screen "P_Slider_1" 1024x768
   Slider "Default" at 10,10 size 60x160; Caption 'SIMATIC'
   TextField "Label_Default" at 10,172 size 68x16; Text 'Default'
   Slider "BackColor" at 80,10 size 60x160; Caption 'SIMATIC'
   TextField "Label_BackColor" at 80,172 size 68x16; Text 'BackColor'
   Slider "BackFillStyle" at 150,10 size 60x160; Caption 'SIMATIC'
   TextField "Label_BackFillStyle" at 150,172 size 68x16; Text 'BackFillStyle'
   Slider "BarBackColor" at 220,10 size 60x160; Caption 'SIMATIC'
   TextField "Label_BarBackColor" at 220,172 size 68x16; Text 'BarBackColor'
   Slider "BarColor" at 290,10 size 60x160; Caption 'SIMATIC'
   TextField "Label_BarColor" at 290,172 size 68x16; Text 'BarColor'
   Slider "BarOrientation" at 360,10 size 60x160; Caption 'SIMATIC'
   TextField "Label_BarOrientation" at 360,172 size 68x16; Text 'BarOrientation'
   Slider "BarOrientation_2" at 430,10 size 60x160; Caption 'SIMATIC'
   TextField "Label_BarOrientation_2" at 430,172 size 68x16; Text 'BarOrientation_2'
   Slider "BarOrientation_3" at 500,10 size 60x160; Caption 'SIMATIC'
   TextField "Label_BarOrientation_3" at 500,172 size 68x16; Text 'BarOrientation_3'
   Slider "BorderBackColor" at 570,10 size 60x160; Caption 'SIMATIC'
   TextField "Label_BorderBackColor" at 570,172 size 68x16; Text 'BorderBackColor'
   Slider "BorderBrightColor3D" at 640,10 size 60x160; Caption 'SIMATIC'
   TextField "Label_BorderBrightColor3D" at 640,172 size 68x16; Text 'BorderBrightColor3D'
   Slider "BorderColor" at 710,10 size 60x160; Caption 'SIMATIC'
   TextField "Label_BorderColor" at 710,172 size 68x16; Text 'BorderColor'
   Slider "BorderInnerStyle3D" at 780,10 size 60x160; Caption 'SIMATIC'
   TextField "Label_BorderInnerStyle3D" at 780,172 size 68x16; Text 'BorderInnerStyle3D'
   Slider "BorderInnerStyle3D_2" at 850,10 size 60x160; Caption 'SIMATIC'
   TextField "Label_BorderInnerStyle3D_2" at 850,172 size 68x16; Text 'BorderInnerStyle3D_2'
   Slider "BorderInnerWidth3D" at 920,10 size 60x160; Caption 'SIMATIC'
   TextField "Label_BorderInnerWidth3D" at 920,172 size 68x16; Text 'BorderInnerWidth3D'
   Slider "BorderOuterStyle3D" at 10,196 size 60x160; Caption 'SIMATIC'
   TextField "Label_BorderOuterStyle3D" at 10,358 size 68x16; Text 'BorderOuterStyle3D'
   Slider "BorderOuterStyle3D_2" at 80,196 size 60x160; Caption 'SIMATIC'
   TextField "Label_BorderOuterStyle3D_2" at 80,358 size 68x16; Text 'BorderOuterStyle3D_2'
   Slider "BorderOuterWidth3D" at 150,196 size 60x160; Caption 'SIMATIC'
   TextField "Label_BorderOuterWidth3D" at 150,358 size 68x16; Text 'BorderOuterWidth3D'
   Slider "BorderShadeColor3D" at 220,196 size 60x160; Caption 'SIMATIC'
   TextField "Label_BorderShadeColor3D" at 220,358 size 68x16; Text 'BorderShadeColor3D'
   Slider "BorderWidth" at 290,196 size 60x160; Caption 'SIMATIC'
   TextField "Label_BorderWidth" at 290,358 size 68x16; Text 'BorderWidth'
   Slider "CornerRadius" at 360,196 size 60x160; Caption 'SIMATIC'
   TextField "Label_CornerRadius" at 360,358 size 68x16; Text 'CornerRadius'
   Slider "EdgeStyle" at 430,196 size 60x160; Caption 'SIMATIC'
   TextField "Label_EdgeStyle" at 430,358 size 68x16; Text 'EdgeStyle'
   Slider "EdgeStyle_2" at 500,196 size 60x160; Caption 'SIMATIC'
   TextField "Label_EdgeStyle_2" at 500,358 size 68x16; Text 'EdgeStyle_2'
   Slider "EdgeStyle_3" at 570,196 size 60x160; Caption 'SIMATIC'
   TextField "Label_EdgeStyle_3" at 570,358 size 68x16; Text 'EdgeStyle_3'
   Slider "EdgeStyle_4" at 640,196 size 60x160; Caption 'SIMATIC'
   TextField "Label_EdgeStyle_4" at 640,358 size 68x16; Text 'EdgeStyle_4'
   Slider "Flashing" at 710,196 size 60x160; Caption 'SIMATIC'
   TextField "Label_Flashing" at 710,358 size 68x16; Text 'Flashing'
   Slider "FocusColor" at 780,196 size 60x160; Caption 'SIMATIC'
   TextField "Label_FocusColor" at 780,358 size 68x16; Text 'FocusColor'
   Slider "FocusWidth" at 850,196 size 60x160; Caption 'SIMATIC'
   TextField "Label_FocusWidth" at 850,358 size 68x16; Text 'FocusWidth'
   Slider "ForeColor" at 920,196 size 60x160; Caption 'SIMATIC'
   TextField "Label_ForeColor" at 920,358 size 68x16; Text 'ForeColor'
   Slider "LabelColor" at 10,382 size 60x160; Caption 'SIMATIC'
   TextField "Label_LabelColor" at 10,544 size 68x16; Text 'LabelColor'
   Slider "MaximumValue" at 80,382 size 60x160; Caption 'SIMATIC'
   TextField "Label_MaximumValue" at 80,544 size 68x16; Text 'MaximumValue'
   Slider "MinimumValue" at 150,382 size 60x160; Caption 'SIMATIC'
   TextField "Label_MinimumValue" at 150,544 size 68x16; Text 'MinimumValue'
   Slider "RangeLower1Color" at 220,382 size 60x160; Caption 'SIMATIC'
   TextField "Label_RangeLower1Color" at 220,544 size 68x16; Text 'RangeLower1Color'
   Slider "RangeLower1Enabled" at 290,382 size 60x160; Caption 'SIMATIC'
   TextField "Label_RangeLower1Enabled" at 290,544 size 68x16; Text 'RangeLower1Enabled'
   Slider "RangeLower2Color" at 360,382 size 60x160; Caption 'SIMATIC'
   TextField "Label_RangeLower2Color" at 360,544 size 68x16; Text 'RangeLower2Color'
   Slider "RangeLower2Enabled" at 430,382 size 60x160; Caption 'SIMATIC'
   TextField "Label_RangeLower2Enabled" at 430,544 size 68x16; Text 'RangeLower2Enabled'
   Slider "RangeNormalColor" at 500,382 size 60x160; Caption 'SIMATIC'
   TextField "Label_RangeNormalColor" at 500,544 size 68x16; Text 'RangeNormalColor'
   Slider "RangeNormalEnabled" at 570,382 size 60x160; Caption 'SIMATIC'
   TextField "Label_RangeNormalEnabled" at 570,544 size 68x16; Text 'RangeNormalEnabled'
   Slider "RangeUpper1Color" at 640,382 size 60x160; Caption 'SIMATIC'
   TextField "Label_RangeUpper1Color" at 640,544 size 68x16; Text 'RangeUpper1Color'
   Slider "RangeUpper1Enabled" at 710,382 size 60x160; Caption 'SIMATIC'
   TextField "Label_RangeUpper1Enabled" at 710,544 size 68x16; Text 'RangeUpper1Enabled'
   Slider "RangeUpper2Color" at 780,382 size 60x160; Caption 'SIMATIC'
   TextField "Label_RangeUpper2Color" at 780,544 size 68x16; Text 'RangeUpper2Color'
   Slider "RangeUpper2Enabled" at 850,382 size 60x160; Caption 'SIMATIC'
   TextField "Label_RangeUpper2Enabled" at 850,544 size 68x16; Text 'RangeUpper2Enabled'
   Slider "ScalePosition" at 920,382 size 60x160; Caption 'SIMATIC'
   TextField "Label_ScalePosition" at 920,544 size 68x16; Text 'ScalePosition'
   Button "Next" at 982,744 size 40x22; TextOff 'Text'
      on Click: ActivateScreen("P_Slider_2", 0)

screen "P_Slider_2" 1024x768
   Slider "ShowBar" at 10,10 size 60x160; Caption 'SIMATIC'
   TextField "Label_ShowBar" at 10,172 size 68x16; Text 'ShowBar'
   Slider "ShowLimitLines" at 80,10 size 60x160; Caption 'SIMATIC'
   TextField "Label_ShowLimitLines" at 80,172 size 68x16; Text 'ShowLimitLines'
   Slider "ShowLimitMarkers" at 150,10 size 60x160; Caption 'SIMATIC'
   TextField "Label_ShowLimitMarkers" at 150,172 size 68x16; Text 'ShowLimitMarkers'
   Slider "ShowLimitRanges" at 220,10 size 60x160; Caption 'SIMATIC'
   TextField "Label_ShowLimitRanges" at 220,172 size 68x16; Text 'ShowLimitRanges'
   Slider "ShowPosition" at 290,10 size 60x160; Caption 'SIMATIC'
   TextField "Label_ShowPosition" at 290,172 size 68x16; Text 'ShowPosition'
   Slider "ShowScale" at 360,10 size 60x160; Caption 'SIMATIC'
   TextField "Label_ShowScale" at 360,172 size 68x16; Text 'ShowScale'
   Slider "ShowThumb" at 430,10 size 60x160; Caption 'SIMATIC'
   TextField "Label_ShowThumb" at 430,172 size 68x16; Text 'ShowThumb'
   Slider "ShowTickLabels" at 500,10 size 60x160; Caption 'SIMATIC'
   TextField "Label_ShowTickLabels" at 500,172 size 68x16; Text 'ShowTickLabels'
   Slider "ShowTicks" at 570,10 size 60x160; Caption 'SIMATIC'
   TextField "Label_ShowTicks" at 570,172 size 68x16; Text 'ShowTicks'
   Slider "ThumbBackColor" at 640,10 size 60x160; Caption 'SIMATIC'
   TextField "Label_ThumbBackColor" at 640,172 size 68x16; Text 'ThumbBackColor'
   Slider "UseDesignColorSchema" at 710,10 size 60x160; Caption 'SIMATIC'
   TextField "Label_UseDesignColorSchema" at 710,172 size 68x16; Text 'UseDesignColorSchema'
   Button "Next" at 982,744 size 40x22; TextOff 'Text'
      on Click: ActivateScreen("P_Gauge_1", 0)

screen "P_Gauge_1" 1024x768
   Gauge "Default" at 10,10 size 150x150; CaptionText 'SIMATIC'
   TextField "Label_Default" at 10,162 size 158x16; Text 'Default'
   Gauge "AngleMax" at 170,10 size 150x150; CaptionText 'SIMATIC'
   TextField "Label_AngleMax" at 170,162 size 158x16; Text 'AngleMax'
   Gauge "AngleMin" at 330,10 size 150x150; CaptionText 'SIMATIC'
   TextField "Label_AngleMin" at 330,162 size 158x16; Text 'AngleMin'
   Gauge "BackColor" at 490,10 size 150x150; CaptionText 'SIMATIC'
   TextField "Label_BackColor" at 490,162 size 158x16; Text 'BackColor'
   Gauge "BackFillStyle" at 650,10 size 150x150; CaptionText 'SIMATIC'
   TextField "Label_BackFillStyle" at 650,162 size 158x16; Text 'BackFillStyle'
   Gauge "BorderBackColor" at 810,10 size 150x150; CaptionText 'SIMATIC'
   TextField "Label_BorderBackColor" at 810,162 size 158x16; Text 'BorderBackColor'
   Gauge "BorderColor" at 10,186 size 150x150; CaptionText 'SIMATIC'
   TextField "Label_BorderColor" at 10,338 size 158x16; Text 'BorderColor'
   Gauge "BorderWidth" at 170,186 size 150x150; CaptionText 'SIMATIC'
   TextField "Label_BorderWidth" at 170,338 size 158x16; Text 'BorderWidth'
   Gauge "CaptionColor" at 330,186 size 150x150; CaptionText 'SIMATIC'
   TextField "Label_CaptionColor" at 330,338 size 158x16; Text 'CaptionColor'
   Gauge "CaptionTop" at 490,186 size 150x150; CaptionText 'SIMATIC'
   TextField "Label_CaptionTop" at 490,338 size 158x16; Text 'CaptionTop'
   Gauge "CenterColor" at 650,186 size 150x150; CaptionText 'SIMATIC'
   TextField "Label_CenterColor" at 650,338 size 158x16; Text 'CenterColor'
   Gauge "CenterSize" at 810,186 size 150x150; CaptionText 'SIMATIC'
   TextField "Label_CenterSize" at 810,338 size 158x16; Text 'CenterSize'
   Gauge "CornerRadius" at 10,362 size 150x150; CaptionText 'SIMATIC'
   TextField "Label_CornerRadius" at 10,514 size 158x16; Text 'CornerRadius'
   Gauge "DialColor" at 170,362 size 150x150; CaptionText 'SIMATIC'
   TextField "Label_DialColor" at 170,514 size 158x16; Text 'DialColor'
   Gauge "DialFillStyle" at 330,362 size 150x150; CaptionText 'SIMATIC'
   TextField "Label_DialFillStyle" at 330,514 size 158x16; Text 'DialFillStyle'
   Gauge "DialSize" at 490,362 size 150x150; CaptionText 'SIMATIC'
   TextField "Label_DialSize" at 490,514 size 158x16; Text 'DialSize'
   Gauge "EdgeStyle" at 650,362 size 150x150; CaptionText 'SIMATIC'
   TextField "Label_EdgeStyle" at 650,514 size 158x16; Text 'EdgeStyle'
   Gauge "EdgeStyle_2" at 810,362 size 150x150; CaptionText 'SIMATIC'
   TextField "Label_EdgeStyle_2" at 810,514 size 158x16; Text 'EdgeStyle_2'
   Gauge "EdgeStyle_3" at 10,538 size 150x150; CaptionText 'SIMATIC'
   TextField "Label_EdgeStyle_3" at 10,690 size 158x16; Text 'EdgeStyle_3'
   Gauge "EdgeStyle_4" at 170,538 size 150x150; CaptionText 'SIMATIC'
   TextField "Label_EdgeStyle_4" at 170,690 size 158x16; Text 'EdgeStyle_4'
   Gauge "Gradation" at 330,538 size 150x150; CaptionText 'SIMATIC'
   TextField "Label_Gradation" at 330,690 size 158x16; Text 'Gradation'
   Gauge "InnerDialColor" at 490,538 size 150x150; CaptionText 'SIMATIC'
   TextField "Label_InnerDialColor" at 490,690 size 158x16; Text 'InnerDialColor'
   Gauge "InnerDialInnerDistance" at 650,538 size 150x150; CaptionText 'SIMATIC'
   TextField "Label_InnerDialInnerDistance" at 650,690 size 158x16; Text 'InnerDialInnerDistance'
   Gauge "InnerDialOuterDistance" at 810,538 size 150x150; CaptionText 'SIMATIC'
   TextField "Label_InnerDialOuterDistance" at 810,690 size 158x16; Text 'InnerDialOuterDistance'
   Button "Next" at 982,744 size 40x22; TextOff 'Text'
      on Click: ActivateScreen("P_Gauge_2", 0)

screen "P_Gauge_2" 1024x768
   Gauge "LockSquaredExtent" at 10,10 size 150x150; CaptionText 'SIMATIC'
   TextField "Label_LockSquaredExtent" at 10,162 size 158x16; Text 'LockSquaredExtent'
   Gauge "MaximumValue" at 170,10 size 150x150; CaptionText 'SIMATIC'
   TextField "Label_MaximumValue" at 170,162 size 158x16; Text 'MaximumValue'
   Gauge "MinimumValue" at 330,10 size 150x150; CaptionText 'SIMATIC'
   TextField "Label_MinimumValue" at 330,162 size 158x16; Text 'MinimumValue'
   Gauge "NeedleHeight" at 490,10 size 150x150; CaptionText 'SIMATIC'
   TextField "Label_NeedleHeight" at 490,162 size 158x16; Text 'NeedleHeight'
   Gauge "PointerColor" at 650,10 size 150x150; CaptionText 'SIMATIC'
   TextField "Label_PointerColor" at 650,162 size 158x16; Text 'PointerColor'
   Gauge "RangeLower1Color" at 810,10 size 150x150; CaptionText 'SIMATIC'
   TextField "Label_RangeLower1Color" at 810,162 size 158x16; Text 'RangeLower1Color'
   Gauge "RangeLower1Enabled" at 10,186 size 150x150; CaptionText 'SIMATIC'
   TextField "Label_RangeLower1Enabled" at 10,338 size 158x16; Text 'RangeLower1Enabled'
   Gauge "RangeLower2Color" at 170,186 size 150x150; CaptionText 'SIMATIC'
   TextField "Label_RangeLower2Color" at 170,338 size 158x16; Text 'RangeLower2Color'
   Gauge "RangeLower2Enabled" at 330,186 size 150x150; CaptionText 'SIMATIC'
   TextField "Label_RangeLower2Enabled" at 330,338 size 158x16; Text 'RangeLower2Enabled'
   Gauge "RangeNormalColor" at 490,186 size 150x150; CaptionText 'SIMATIC'
   TextField "Label_RangeNormalColor" at 490,338 size 158x16; Text 'RangeNormalColor'
   Gauge "RangeNormalEnabled" at 650,186 size 150x150; CaptionText 'SIMATIC'
   TextField "Label_RangeNormalEnabled" at 650,338 size 158x16; Text 'RangeNormalEnabled'
   Gauge "RangeUpper1Color" at 810,186 size 150x150; CaptionText 'SIMATIC'
   TextField "Label_RangeUpper1Color" at 810,338 size 158x16; Text 'RangeUpper1Color'
   Gauge "RangeUpper1Enabled" at 10,362 size 150x150; CaptionText 'SIMATIC'
   TextField "Label_RangeUpper1Enabled" at 10,514 size 158x16; Text 'RangeUpper1Enabled'
   Gauge "RangeUpper1Start" at 170,362 size 150x150; CaptionText 'SIMATIC'
   TextField "Label_RangeUpper1Start" at 170,514 size 158x16; Text 'RangeUpper1Start'
   Gauge "RangeUpper2Color" at 330,362 size 150x150; CaptionText 'SIMATIC'
   TextField "Label_RangeUpper2Color" at 330,514 size 158x16; Text 'RangeUpper2Color'
   Gauge "RangeUpper2Enabled" at 490,362 size 150x150; CaptionText 'SIMATIC'
   TextField "Label_RangeUpper2Enabled" at 490,514 size 158x16; Text 'RangeUpper2Enabled'
   Gauge "RangeUpper2Start" at 650,362 size 150x150; CaptionText 'SIMATIC'
   TextField "Label_RangeUpper2Start" at 650,514 size 158x16; Text 'RangeUpper2Start'
   Gauge "ScaleLabelColor" at 810,362 size 150x150; CaptionText 'SIMATIC'
   TextField "Label_ScaleLabelColor" at 810,514 size 158x16; Text 'ScaleLabelColor'
   Gauge "ScaleTickColor" at 10,538 size 150x150; CaptionText 'SIMATIC'
   TextField "Label_ScaleTickColor" at 10,690 size 158x16; Text 'ScaleTickColor'
   Gauge "ScaleTickLabelPosition" at 170,538 size 150x150; CaptionText 'SIMATIC'
   TextField "Label_ScaleTickLabelPosition" at 170,690 size 158x16; Text 'ScaleTickLabelPosition'
   Gauge "ScaleTickLength" at 330,538 size 150x150; CaptionText 'SIMATIC'
   TextField "Label_ScaleTickLength" at 330,690 size 158x16; Text 'ScaleTickLength'
   Gauge "ScaleTickPosition" at 490,538 size 150x150; CaptionText 'SIMATIC'
   TextField "Label_ScaleTickPosition" at 490,690 size 158x16; Text 'ScaleTickPosition'
   Gauge "ShowDecimalPoint" at 650,538 size 150x150; CaptionText 'SIMATIC'
   TextField "Label_ShowDecimalPoint" at 650,690 size 158x16; Text 'ShowDecimalPoint'
   Gauge "ShowInnerDial" at 810,538 size 150x150; CaptionText 'SIMATIC'
   TextField "Label_ShowInnerDial" at 810,690 size 158x16; Text 'ShowInnerDial'
   Button "Next" at 982,744 size 40x22; TextOff 'Text'
      on Click: ActivateScreen("P_Gauge_3", 0)

screen "P_Gauge_3" 1024x768
   Gauge "ShowLimitRanges" at 10,10 size 150x150; CaptionText 'SIMATIC'
   TextField "Label_ShowLimitRanges" at 10,162 size 158x16; Text 'ShowLimitRanges'
   Gauge "ShowPeakValuePointer" at 170,10 size 150x150; CaptionText 'SIMATIC'
   TextField "Label_ShowPeakValuePointer" at 170,162 size 158x16; Text 'ShowPeakValuePointer'
   Gauge "UnitColor" at 330,10 size 150x150; CaptionText 'SIMATIC'
   TextField "Label_UnitColor" at 330,162 size 158x16; Text 'UnitColor'
   Gauge "UnitTop" at 490,10 size 150x150; CaptionText 'SIMATIC'
   TextField "Label_UnitTop" at 490,162 size 158x16; Text 'UnitTop'
   Gauge "UseDesignColorSchema" at 650,10 size 150x150; CaptionText 'SIMATIC'
   TextField "Label_UseDesignColorSchema" at 650,162 size 158x16; Text 'UseDesignColorSchema'
   Button "Next" at 982,744 size 40x22; TextOff 'Text'
      on Click: ActivateScreen("P_Clock_1", 0)

screen "P_Clock_1" 1024x768
   Clock "Default" at 10,10 size 150x150
   TextField "Label_Default" at 10,162 size 158x16; Text 'Default'
   Clock "Analog" at 170,10 size 150x150
   TextField "Label_Analog" at 170,162 size 158x16; Text 'Analog'
   Clock "BackFillStyle" at 330,10 size 150x150
   TextField "Label_BackFillStyle" at 330,162 size 158x16; Text 'BackFillStyle'
   Clock "BorderBackColor" at 490,10 size 150x150
   TextField "Label_BorderBackColor" at 490,162 size 158x16; Text 'BorderBackColor'
   Clock "BorderColor" at 650,10 size 150x150
   TextField "Label_BorderColor" at 650,162 size 158x16; Text 'BorderColor'
   Clock "BorderWidth" at 810,10 size 150x150
   TextField "Label_BorderWidth" at 810,162 size 158x16; Text 'BorderWidth'
   Clock "CornerRadius" at 10,186 size 150x150
   TextField "Label_CornerRadius" at 10,338 size 158x16; Text 'CornerRadius'
   Clock "DialColor" at 170,186 size 150x150
   TextField "Label_DialColor" at 170,338 size 158x16; Text 'DialColor'
   Clock "EdgeStyle" at 330,186 size 150x150
   TextField "Label_EdgeStyle" at 330,338 size 158x16; Text 'EdgeStyle'
   Clock "EdgeStyle_2" at 490,186 size 150x150
   TextField "Label_EdgeStyle_2" at 490,338 size 158x16; Text 'EdgeStyle_2'
   Clock "EdgeStyle_3" at 650,186 size 150x150
   TextField "Label_EdgeStyle_3" at 650,338 size 158x16; Text 'EdgeStyle_3'
   Clock "EdgeStyle_4" at 810,186 size 150x150
   TextField "Label_EdgeStyle_4" at 810,338 size 158x16; Text 'EdgeStyle_4'
   Clock "Flashing" at 10,362 size 150x150
   TextField "Label_Flashing" at 10,514 size 158x16; Text 'Flashing'
   Clock "HourNeedleHeight" at 170,362 size 150x150
   TextField "Label_HourNeedleHeight" at 170,514 size 158x16; Text 'HourNeedleHeight'
   Clock "HourNeedleWidth" at 330,362 size 150x150
   TextField "Label_HourNeedleWidth" at 330,514 size 158x16; Text 'HourNeedleWidth'
   Clock "LockSquaredExtent" at 490,362 size 150x150
   TextField "Label_LockSquaredExtent" at 490,514 size 158x16; Text 'LockSquaredExtent'
   Clock "MinuteNeedleHeight" at 650,362 size 150x150
   TextField "Label_MinuteNeedleHeight" at 650,514 size 158x16; Text 'MinuteNeedleHeight'
   Clock "MinuteNeedleWidth" at 810,362 size 150x150
   TextField "Label_MinuteNeedleWidth" at 810,514 size 158x16; Text 'MinuteNeedleWidth'
   Clock "NeedleBorderColor" at 10,538 size 150x150
   TextField "Label_NeedleBorderColor" at 10,690 size 158x16; Text 'NeedleBorderColor'
   Clock "NeedleColor" at 170,538 size 150x150
   TextField "Label_NeedleColor" at 170,690 size 158x16; Text 'NeedleColor'
   Clock "NeedleFillStyle" at 330,538 size 150x150
   TextField "Label_NeedleFillStyle" at 330,690 size 158x16; Text 'NeedleFillStyle'
   Clock "NumberStyle" at 490,538 size 150x150
   TextField "Label_NumberStyle" at 490,690 size 158x16; Text 'NumberStyle'
   Clock "NumberStyle_2" at 650,538 size 150x150
   TextField "Label_NumberStyle_2" at 650,690 size 158x16; Text 'NumberStyle_2'
   Clock "SecondNeedleHeight" at 810,538 size 150x150
   TextField "Label_SecondNeedleHeight" at 810,690 size 158x16; Text 'SecondNeedleHeight'
   Button "Next" at 982,744 size 40x22; TextOff 'Text'
      on Click: ActivateScreen("P_Clock_2", 0)

screen "P_Clock_2" 1024x768
   Clock "SecondNeedleWidth" at 10,10 size 150x150
   TextField "Label_SecondNeedleWidth" at 10,162 size 158x16; Text 'SecondNeedleWidth'
   Clock "ShowTicks" at 170,10 size 150x150
   TextField "Label_ShowTicks" at 170,162 size 158x16; Text 'ShowTicks'
   Clock "TickDistance" at 330,10 size 150x150
   TextField "Label_TickDistance" at 330,162 size 158x16; Text 'TickDistance'
   Clock "TickStyle" at 490,10 size 150x150
   TextField "Label_TickStyle" at 490,162 size 158x16; Text 'TickStyle'
   Clock "TicksColor" at 650,10 size 150x150
   TextField "Label_TicksColor" at 650,162 size 158x16; Text 'TicksColor'
   Clock "UseDesignColorSchema" at 810,10 size 150x150
   TextField "Label_UseDesignColorSchema" at 810,162 size 158x16; Text 'UseDesignColorSchema'
   Button "Next" at 982,744 size 40x22; TextOff 'Text'
      on Click: ActivateScreen("P_Line_1", 0)

screen "P_IOField_1" 1024x768
   IOField "Default" at 10,10 size 100x30
   TextField "Label_Default" at 10,42 size 108x16; Text 'Default'
   IOField "AboveUpperLimitColor" at 120,10 size 100x30
   TextField "Label_AboveUpperLimitColor" at 120,42 size 108x16; Text 'AboveUpperLimitColor'
   IOField "BackColor" at 230,10 size 100x30
   TextField "Label_BackColor" at 230,42 size 108x16; Text 'BackColor'
   IOField "BackFillStyle" at 340,10 size 100x30
   TextField "Label_BackFillStyle" at 340,42 size 108x16; Text 'BackFillStyle'
   IOField "BelowLowerLimitColor" at 450,10 size 100x30
   TextField "Label_BelowLowerLimitColor" at 450,42 size 108x16; Text 'BelowLowerLimitColor'
   IOField "BorderBackColor" at 560,10 size 100x30
   TextField "Label_BorderBackColor" at 560,42 size 108x16; Text 'BorderBackColor'
   IOField "BorderColor" at 670,10 size 100x30
   TextField "Label_BorderColor" at 670,42 size 108x16; Text 'BorderColor'
   IOField "BorderWidth" at 780,10 size 100x30
   TextField "Label_BorderWidth" at 780,42 size 108x16; Text 'BorderWidth'
   IOField "BottomMargin" at 890,10 size 100x30
   TextField "Label_BottomMargin" at 890,42 size 108x16; Text 'BottomMargin'
   IOField "CornerRadius" at 10,66 size 100x30
   TextField "Label_CornerRadius" at 10,98 size 108x16; Text 'CornerRadius'
   IOField "DataFormat_3" at 120,66 size 100x30
   TextField "Label_DataFormat_3" at 120,98 size 108x16; Text 'DataFormat_3'
   IOField "EdgeStyle" at 230,66 size 100x30
   TextField "Label_EdgeStyle" at 230,98 size 108x16; Text 'EdgeStyle'
   IOField "EdgeStyle_2" at 340,66 size 100x30
   TextField "Label_EdgeStyle_2" at 340,98 size 108x16; Text 'EdgeStyle_2'
   IOField "EdgeStyle_3" at 450,66 size 100x30
   TextField "Label_EdgeStyle_3" at 450,98 size 108x16; Text 'EdgeStyle_3'
   IOField "EdgeStyle_4" at 560,66 size 100x30
   TextField "Label_EdgeStyle_4" at 560,98 size 108x16; Text 'EdgeStyle_4'
   IOField "FieldLength" at 670,66 size 100x30
   TextField "Label_FieldLength" at 670,98 size 108x16; Text 'FieldLength'
   IOField "FitToLargest" at 780,66 size 100x30
   TextField "Label_FitToLargest" at 780,98 size 108x16; Text 'FitToLargest'
   IOField "Flashing" at 890,66 size 100x30
   TextField "Label_Flashing" at 890,98 size 108x16; Text 'Flashing'
   IOField "ForeColor" at 10,122 size 100x30
   TextField "Label_ForeColor" at 10,154 size 108x16; Text 'ForeColor'
   IOField "FormatPattern" at 120,122 size 100x30; FormatPattern 99.9
   TextField "Label_FormatPattern" at 120,154 size 108x16; Text 'FormatPattern'
   IOField "HorizontalAlignment" at 230,122 size 100x30
   TextField "Label_HorizontalAlignment" at 230,154 size 108x16; Text 'HorizontalAlignment'
   IOField "HorizontalAlignment_2" at 340,122 size 100x30
   TextField "Label_HorizontalAlignment_2" at 340,154 size 108x16; Text 'HorizontalAlignment_2'
   IOField "LeftMargin" at 450,122 size 100x30
   TextField "Label_LeftMargin" at 450,154 size 108x16; Text 'LeftMargin'
   IOField "Mode" at 560,122 size 100x30
   TextField "Label_Mode" at 560,154 size 108x16; Text 'Mode'
   IOField "Mode_2" at 670,122 size 100x30
   TextField "Label_Mode_2" at 670,154 size 108x16; Text 'Mode_2'
   IOField "RightMargin" at 780,122 size 100x30
   TextField "Label_RightMargin" at 780,154 size 108x16; Text 'RightMargin'
   IOField "ShiftDecimalPoint" at 890,122 size 100x30
   TextField "Label_ShiftDecimalPoint" at 890,154 size 108x16; Text 'ShiftDecimalPoint'
   IOField "ShowLeadingZeros" at 10,178 size 100x30
   TextField "Label_ShowLeadingZeros" at 10,210 size 108x16; Text 'ShowLeadingZeros'
   IOField "TopMargin" at 120,178 size 100x30
   TextField "Label_TopMargin" at 120,210 size 108x16; Text 'TopMargin'
   IOField "Unit" at 230,178 size 100x30; Unit mm
   TextField "Label_Unit" at 230,210 size 108x16; Text 'Unit'
   IOField "UseDesignColorSchema" at 340,178 size 100x30
   TextField "Label_UseDesignColorSchema" at 340,210 size 108x16; Text 'UseDesignColorSchema'
   IOField "VerticalAlignment" at 450,178 size 100x30
   TextField "Label_VerticalAlignment" at 450,210 size 108x16; Text 'VerticalAlignment'
   IOField "VerticalAlignment_2" at 560,178 size 100x30
   TextField "Label_VerticalAlignment_2" at 560,210 size 108x16; Text 'VerticalAlignment_2'
   Button "Next" at 982,744 size 40x22; TextOff 'Text'
      on Click: ActivateScreen("P_Button_1", 0)

screen "D_Bar_1" 1024x768
   Bar "Static" at 6,4 size 40x120
   TextField "Label_Static" at 6,156 size 88x16; Text 'Static'
   Bar "A_Range" at 98,4 size 40x120
      Appearance <- "D_Range"
   TextField "Label_A_Range" at 98,156 size 88x16; Text 'A_Range'
   Bar "A_Flash" at 190,4 size 40x120
      Appearance <- "D_Range"
   TextField "Label_A_Flash" at 190,156 size 88x16; Text 'A_Flash'
   Bar "A_Bit" at 282,4 size 40x120
      Appearance <- "D_Bool"
   TextField "Label_A_Bit" at 282,156 size 88x16; Text 'A_Bit'
   Bar "A_Bits" at 374,4 size 40x120
      Appearance <- "D_Bits"
   TextField "Label_A_Bits" at 374,156 size 88x16; Text 'A_Bits'
   Bar "V_Range" at 466,4 size 40x120
      Visibility <- "D_Range"
   TextField "Label_V_Range" at 466,156 size 88x16; Text 'V_Range'
   Bar "V_Bit" at 558,4 size 40x120
      Visibility <- "D_Vis"
   TextField "Label_V_Bit" at 558,156 size 88x16; Text 'V_Bit'
   Bar "M_H" at 650,4 size 40x120
      HorizontalMovement <- "D_Pct"
   TextField "Label_M_H" at 650,156 size 88x16; Text 'M_H'
   Bar "M_V" at 742,4 size 40x120
      VerticalMovement <- "D_Pct"
   TextField "Label_M_V" at 742,156 size 88x16; Text 'M_V'
   Bar "M_D" at 834,4 size 40x120
      DiagonalMovement <- "D_Pct"
   TextField "Label_M_D" at 834,156 size 88x16; Text 'M_D'
   Bar "M_Direct" at 926,4 size 40x120
      DirectMovement <- "D_X"
      DirectMovement <- "D_Y"
   TextField "Label_M_Direct" at 926,156 size 88x16; Text 'M_Direct'
   Bar "E_Range" at 6,176 size 40x120
      ObjectEnable <- "D_Range"
   TextField "Label_E_Range" at 6,328 size 88x16; Text 'E_Range'
   Bar "E_Bit" at 98,176 size 40x120
      ObjectEnable <- "D_En"
   TextField "Label_E_Bit" at 98,328 size 88x16; Text 'E_Bit'
   Bar "PV_Pct" at 190,176 size 40x120
      ProcessValue <- "D_Pct"
   TextField "Label_PV_Pct" at 190,328 size 88x16; Text 'PV_Pct'
   Bar "PV_Real" at 282,176 size 40x120
      ProcessValue <- "D_Real"
   TextField "Label_PV_Real" at 282,328 size 88x16; Text 'PV_Real'
   Bar "PV_BarR" at 374,176 size 40x120
      ProcessValue <- "D_BarR"
   TextField "Label_PV_BarR" at 374,328 size 88x16; Text 'PV_BarR'
   Bar "PV_Pct_0_100" at 466,176 size 40x120; MinimumValue 0; MaximumValue 100
      ProcessValue <- "D_Pct"
   TextField "Label_PV_Pct_0_100" at 466,328 size 88x16; Text 'PV_Pct_0_100'
   Bar "PV_Pct_MaxMin" at 558,176 size 40x120
      ProcessValue <- "D_Pct"
      MaximumValue <- "D_Max"
      MinimumValue <- "D_Min"
   TextField "Label_PV_Pct_MaxMin" at 558,328 size 88x16; Text 'PV_Pct_MaxMin'
   IOField "State" at 4,742 size 60x22; FormatPattern 9
      ProcessValue <- "D_State"
   Button "S1" at 70,742 size 40x22; TextOff 'S1'
      on Click: "SetS1"()
   Button "S2" at 114,742 size 40x22; TextOff 'S2'
      on Click: "SetS2"()
   Button "S3" at 158,742 size 40x22; TextOff 'S3'
      on Click: "SetS3"()
   Button "S4" at 202,742 size 40x22; TextOff 'S4'
      on Click: "SetS4"()
   Button "Next" at 980,742 size 40x22; TextOff 'Next'
      on Click: ActivateScreen("D_Switch_1", 0)

screen "D_Button_1" 1024x768
   Button "Static" at 6,4 size 100x40; TextOff 'Text'
   TextField "Label_Static" at 6,76 size 148x16; Text 'Static'
   Button "A_Range" at 158,4 size 100x40; TextOff 'Text'
      Appearance <- "D_Range"
   TextField "Label_A_Range" at 158,76 size 148x16; Text 'A_Range'
   Button "A_Flash" at 310,4 size 100x40; TextOff 'Text'
      Appearance <- "D_Range"
   TextField "Label_A_Flash" at 310,76 size 148x16; Text 'A_Flash'
   Button "A_Bit" at 462,4 size 100x40; TextOff 'Text'
      Appearance <- "D_Bool"
   TextField "Label_A_Bit" at 462,76 size 148x16; Text 'A_Bit'
   Button "A_Bits" at 614,4 size 100x40; TextOff 'Text'
      Appearance <- "D_Bits"
   TextField "Label_A_Bits" at 614,76 size 148x16; Text 'A_Bits'
   Button "V_Range" at 766,4 size 100x40; TextOff 'Text'
      Visibility <- "D_Range"
   TextField "Label_V_Range" at 766,76 size 148x16; Text 'V_Range'
   Button "V_Bit" at 6,96 size 100x40; TextOff 'Text'
      Visibility <- "D_Vis"
   TextField "Label_V_Bit" at 6,168 size 148x16; Text 'V_Bit'
   Button "M_H" at 158,96 size 100x40; TextOff 'Text'
      HorizontalMovement <- "D_Pct"
   TextField "Label_M_H" at 158,168 size 148x16; Text 'M_H'
   Button "M_V" at 310,96 size 100x40; TextOff 'Text'
      VerticalMovement <- "D_Pct"
   TextField "Label_M_V" at 310,168 size 148x16; Text 'M_V'
   Button "M_D" at 462,96 size 100x40; TextOff 'Text'
      DiagonalMovement <- "D_Pct"
   TextField "Label_M_D" at 462,168 size 148x16; Text 'M_D'
   Button "M_Direct" at 614,96 size 100x40; TextOff 'Text'
      DirectMovement <- "D_X"
      DirectMovement <- "D_Y"
   TextField "Label_M_Direct" at 614,168 size 148x16; Text 'M_Direct'
   Button "E_Range" at 766,96 size 100x40; TextOff 'Text'
      ObjectEnable <- "D_Range"
   TextField "Label_E_Range" at 766,168 size 148x16; Text 'E_Range'
   Button "E_Bit" at 6,188 size 100x40; TextOff 'Text'
      ObjectEnable <- "D_En"
   TextField "Label_E_Bit" at 6,260 size 148x16; Text 'E_Bit'
   IOField "State" at 4,742 size 60x22; FormatPattern 9
      ProcessValue <- "D_State"
   Button "S1" at 70,742 size 40x22; TextOff 'S1'
      on Click: "SetS1"()
   Button "S2" at 114,742 size 40x22; TextOff 'S2'
      on Click: "SetS2"()
   Button "S3" at 158,742 size 40x22; TextOff 'S3'
      on Click: "SetS3"()
   Button "S4" at 202,742 size 40x22; TextOff 'S4'
      on Click: "SetS4"()
   Button "Next" at 980,742 size 40x22; TextOff 'Next'
      on Click: ActivateScreen("D_SymbolicIOField_1", 0)

screen "D_Circle_1" 1024x768
   TextField "Label_Static" at 6,86 size 98x16; Text 'Static'
   Circle "A_Range" at 108,4 size 50x50
      Appearance <- "D_Range"
   TextField "Label_A_Range" at 108,86 size 98x16; Text 'A_Range'
   Circle "A_Flash" at 210,4 size 50x50
      Appearance <- "D_Range"
   TextField "Label_A_Flash" at 210,86 size 98x16; Text 'A_Flash'
   Circle "A_Bit" at 312,4 size 50x50
      Appearance <- "D_Bool"
   TextField "Label_A_Bit" at 312,86 size 98x16; Text 'A_Bit'
   Circle "A_Bits" at 414,4 size 50x50
      Appearance <- "D_Bits"
   TextField "Label_A_Bits" at 414,86 size 98x16; Text 'A_Bits'
   Circle "V_Range" at 516,4 size 50x50
      Visibility <- "D_Range"
   TextField "Label_V_Range" at 516,86 size 98x16; Text 'V_Range'
   Circle "V_Bit" at 618,4 size 50x50
      Visibility <- "D_Vis"
   TextField "Label_V_Bit" at 618,86 size 98x16; Text 'V_Bit'
   Circle "M_H" at 720,4 size 50x50
      HorizontalMovement <- "D_Pct"
   TextField "Label_M_H" at 720,86 size 98x16; Text 'M_H'
   Circle "M_V" at 822,4 size 50x50
      VerticalMovement <- "D_Pct"
   TextField "Label_M_V" at 822,86 size 98x16; Text 'M_V'
   Circle "M_D" at 6,106 size 50x50
      DiagonalMovement <- "D_Pct"
   TextField "Label_M_D" at 6,188 size 98x16; Text 'M_D'
   Circle "M_Direct" at 108,106 size 50x50
      DirectMovement <- "D_X"
      DirectMovement <- "D_Y"
   TextField "Label_M_Direct" at 108,188 size 98x16; Text 'M_Direct'
   Circle "E_Range" at 210,106 size 50x50
      ObjectEnable <- "D_Range"
   TextField "Label_E_Range" at 210,188 size 98x16; Text 'E_Range'
   Circle "E_Bit" at 312,106 size 50x50
      ObjectEnable <- "D_En"
   TextField "Label_E_Bit" at 312,188 size 98x16; Text 'E_Bit'
   IOField "State" at 4,742 size 60x22; FormatPattern 9
      ProcessValue <- "D_State"
   Button "S1" at 70,742 size 40x22; TextOff 'S1'
      on Click: "SetS1"()
   Button "S2" at 114,742 size 40x22; TextOff 'S2'
      on Click: "SetS2"()
   Button "S3" at 158,742 size 40x22; TextOff 'S3'
      on Click: "SetS3"()
   Button "S4" at 202,742 size 40x22; TextOff 'S4'
      on Click: "SetS4"()
   Button "Next" at 980,742 size 40x22; TextOff 'Next'
      on Click: ActivateScreen("D_Rectangle_1", 0)

screen "D_Clock_1" 1024x768
   Clock "Static" at 6,4 size 150x150
   TextField "Label_Static" at 6,186 size 198x16; Text 'Static'
   Clock "A_Range" at 208,4 size 150x150
      Appearance <- "D_Range"
   TextField "Label_A_Range" at 208,186 size 198x16; Text 'A_Range'
   Clock "A_Flash" at 410,4 size 150x150
      Appearance <- "D_Range"
   TextField "Label_A_Flash" at 410,186 size 198x16; Text 'A_Flash'
   Clock "A_Bit" at 612,4 size 150x150
      Appearance <- "D_Bool"
   TextField "Label_A_Bit" at 612,186 size 198x16; Text 'A_Bit'
   Clock "A_Bits" at 814,4 size 150x150
      Appearance <- "D_Bits"
   TextField "Label_A_Bits" at 814,186 size 198x16; Text 'A_Bits'
   Clock "V_Range" at 6,206 size 150x150
      Visibility <- "D_Range"
   TextField "Label_V_Range" at 6,388 size 198x16; Text 'V_Range'
   Clock "V_Bit" at 208,206 size 150x150
      Visibility <- "D_Vis"
   TextField "Label_V_Bit" at 208,388 size 198x16; Text 'V_Bit'
   Clock "M_H" at 410,206 size 150x150
      HorizontalMovement <- "D_Pct"
   TextField "Label_M_H" at 410,388 size 198x16; Text 'M_H'
   Clock "M_V" at 612,206 size 150x150
      VerticalMovement <- "D_Pct"
   TextField "Label_M_V" at 612,388 size 198x16; Text 'M_V'
   Clock "M_D" at 814,206 size 150x150
      DiagonalMovement <- "D_Pct"
   TextField "Label_M_D" at 814,388 size 198x16; Text 'M_D'
   Clock "M_Direct" at 6,408 size 150x150
      DirectMovement <- "D_X"
      DirectMovement <- "D_Y"
   TextField "Label_M_Direct" at 6,590 size 198x16; Text 'M_Direct'
   Clock "E_Range" at 208,408 size 150x150
      ObjectEnable <- "D_Range"
   TextField "Label_E_Range" at 208,590 size 198x16; Text 'E_Range'
   Clock "E_Bit" at 410,408 size 150x150
      ObjectEnable <- "D_En"
   TextField "Label_E_Bit" at 410,590 size 198x16; Text 'E_Bit'
   IOField "State" at 4,742 size 60x22; FormatPattern 9
      ProcessValue <- "D_State"
   Button "S1" at 70,742 size 40x22; TextOff 'S1'
      on Click: "SetS1"()
   Button "S2" at 114,742 size 40x22; TextOff 'S2'
      on Click: "SetS2"()
   Button "S3" at 158,742 size 40x22; TextOff 'S3'
      on Click: "SetS3"()
   Button "S4" at 202,742 size 40x22; TextOff 'S4'
      on Click: "SetS4"()
   Button "Next" at 980,742 size 40x22; TextOff 'Next'
      on Click: ActivateScreen("D_Line_1", 0)

screen "D_DateTimeField_1" 1024x768
   DateTimeField "Static" at 6,4 size 160x30
   TextField "Label_Static" at 6,66 size 208x16; Text 'Static'
   DateTimeField "A_Range" at 218,4 size 160x30
      Appearance <- "D_Range"
   TextField "Label_A_Range" at 218,66 size 208x16; Text 'A_Range'
   DateTimeField "A_Flash" at 430,4 size 160x30
      Appearance <- "D_Range"
   TextField "Label_A_Flash" at 430,66 size 208x16; Text 'A_Flash'
   DateTimeField "A_Bit" at 642,4 size 160x30
      Appearance <- "D_Bool"
   TextField "Label_A_Bit" at 642,66 size 208x16; Text 'A_Bit'
   DateTimeField "A_Bits" at 6,86 size 160x30
      Appearance <- "D_Bits"
   TextField "Label_A_Bits" at 6,148 size 208x16; Text 'A_Bits'
   DateTimeField "V_Range" at 218,86 size 160x30
      Visibility <- "D_Range"
   TextField "Label_V_Range" at 218,148 size 208x16; Text 'V_Range'
   DateTimeField "V_Bit" at 430,86 size 160x30
      Visibility <- "D_Vis"
   TextField "Label_V_Bit" at 430,148 size 208x16; Text 'V_Bit'
   DateTimeField "M_H" at 642,86 size 160x30
      HorizontalMovement <- "D_Pct"
   TextField "Label_M_H" at 642,148 size 208x16; Text 'M_H'
   DateTimeField "M_V" at 6,168 size 160x30
      VerticalMovement <- "D_Pct"
   TextField "Label_M_V" at 6,230 size 208x16; Text 'M_V'
   DateTimeField "M_D" at 218,168 size 160x30
      DiagonalMovement <- "D_Pct"
   TextField "Label_M_D" at 218,230 size 208x16; Text 'M_D'
   DateTimeField "M_Direct" at 430,168 size 160x30
      DirectMovement <- "D_X"
      DirectMovement <- "D_Y"
   TextField "Label_M_Direct" at 430,230 size 208x16; Text 'M_Direct'
   DateTimeField "E_Range" at 642,168 size 160x30
      ObjectEnable <- "D_Range"
   TextField "Label_E_Range" at 642,230 size 208x16; Text 'E_Range'
   DateTimeField "E_Bit" at 6,250 size 160x30
      ObjectEnable <- "D_En"
   TextField "Label_E_Bit" at 6,312 size 208x16; Text 'E_Bit'
   DateTimeField "PV_DateTime" at 218,250 size 160x30
      ProcessValue <- "D_DateTime"
   TextField "Label_PV_DateTime" at 218,312 size 208x16; Text 'PV_DateTime'
   IOField "State" at 4,742 size 60x22; FormatPattern 9
      ProcessValue <- "D_State"
   Button "S1" at 70,742 size 40x22; TextOff 'S1'
      on Click: "SetS1"()
   Button "S2" at 114,742 size 40x22; TextOff 'S2'
      on Click: "SetS2"()
   Button "S3" at 158,742 size 40x22; TextOff 'S3'
      on Click: "SetS3"()
   Button "S4" at 202,742 size 40x22; TextOff 'S4'
      on Click: "SetS4"()
   Button "Next" at 980,742 size 40x22; TextOff 'Next'
      on Click: ActivateScreen("D_Bar_1", 0)

screen "D_Ellipse_1" 1024x768
   TextField "Label_Static" at 6,86 size 148x16; Text 'Static'
   Ellipse "A_Range" at 158,4 size 100x50
      Appearance <- "D_Range"
   TextField "Label_A_Range" at 158,86 size 148x16; Text 'A_Range'
   Ellipse "A_Flash" at 310,4 size 100x50
      Appearance <- "D_Range"
   TextField "Label_A_Flash" at 310,86 size 148x16; Text 'A_Flash'
   Ellipse "A_Bit" at 462,4 size 100x50
      Appearance <- "D_Bool"
   TextField "Label_A_Bit" at 462,86 size 148x16; Text 'A_Bit'
   Ellipse "A_Bits" at 614,4 size 100x50
      Appearance <- "D_Bits"
   TextField "Label_A_Bits" at 614,86 size 148x16; Text 'A_Bits'
   Ellipse "V_Range" at 766,4 size 100x50
      Visibility <- "D_Range"
   TextField "Label_V_Range" at 766,86 size 148x16; Text 'V_Range'
   Ellipse "V_Bit" at 6,106 size 100x50
      Visibility <- "D_Vis"
   TextField "Label_V_Bit" at 6,188 size 148x16; Text 'V_Bit'
   Ellipse "M_H" at 158,106 size 100x50
      HorizontalMovement <- "D_Pct"
   TextField "Label_M_H" at 158,188 size 148x16; Text 'M_H'
   Ellipse "M_V" at 310,106 size 100x50
      VerticalMovement <- "D_Pct"
   TextField "Label_M_V" at 310,188 size 148x16; Text 'M_V'
   Ellipse "M_D" at 462,106 size 100x50
      DiagonalMovement <- "D_Pct"
   TextField "Label_M_D" at 462,188 size 148x16; Text 'M_D'
   Ellipse "M_Direct" at 614,106 size 100x50
      DirectMovement <- "D_X"
      DirectMovement <- "D_Y"
   TextField "Label_M_Direct" at 614,188 size 148x16; Text 'M_Direct'
   Ellipse "E_Range" at 766,106 size 100x50
      ObjectEnable <- "D_Range"
   TextField "Label_E_Range" at 766,188 size 148x16; Text 'E_Range'
   Ellipse "E_Bit" at 6,208 size 100x50
      ObjectEnable <- "D_En"
   TextField "Label_E_Bit" at 6,290 size 148x16; Text 'E_Bit'
   IOField "State" at 4,742 size 60x22; FormatPattern 9
      ProcessValue <- "D_State"
   Button "S1" at 70,742 size 40x22; TextOff 'S1'
      on Click: "SetS1"()
   Button "S2" at 114,742 size 40x22; TextOff 'S2'
      on Click: "SetS2"()
   Button "S3" at 158,742 size 40x22; TextOff 'S3'
      on Click: "SetS3"()
   Button "S4" at 202,742 size 40x22; TextOff 'S4'
      on Click: "SetS4"()
   Button "Next" at 980,742 size 40x22; TextOff 'Next'
      on Click: ActivateScreen("D_Circle_1", 0)

screen "D_Gauge_1" 1024x768
   Gauge "Static" at 6,4 size 150x150; CaptionText 'SIMATIC'
   TextField "Label_Static" at 6,186 size 198x16; Text 'Static'
   Gauge "A_Range" at 208,4 size 150x150; CaptionText 'SIMATIC'
      Appearance <- "D_Range"
   TextField "Label_A_Range" at 208,186 size 198x16; Text 'A_Range'
   Gauge "A_Flash" at 410,4 size 150x150; CaptionText 'SIMATIC'
      Appearance <- "D_Range"
   TextField "Label_A_Flash" at 410,186 size 198x16; Text 'A_Flash'
   Gauge "A_Bit" at 612,4 size 150x150; CaptionText 'SIMATIC'
      Appearance <- "D_Bool"
   TextField "Label_A_Bit" at 612,186 size 198x16; Text 'A_Bit'
   Gauge "A_Bits" at 814,4 size 150x150; CaptionText 'SIMATIC'
      Appearance <- "D_Bits"
   TextField "Label_A_Bits" at 814,186 size 198x16; Text 'A_Bits'
   Gauge "V_Range" at 6,206 size 150x150; CaptionText 'SIMATIC'
      Visibility <- "D_Range"
   TextField "Label_V_Range" at 6,388 size 198x16; Text 'V_Range'
   Gauge "V_Bit" at 208,206 size 150x150; CaptionText 'SIMATIC'
      Visibility <- "D_Vis"
   TextField "Label_V_Bit" at 208,388 size 198x16; Text 'V_Bit'
   Gauge "M_H" at 410,206 size 150x150; CaptionText 'SIMATIC'
      HorizontalMovement <- "D_Pct"
   TextField "Label_M_H" at 410,388 size 198x16; Text 'M_H'
   Gauge "M_V" at 612,206 size 150x150; CaptionText 'SIMATIC'
      VerticalMovement <- "D_Pct"
   TextField "Label_M_V" at 612,388 size 198x16; Text 'M_V'
   Gauge "M_D" at 814,206 size 150x150; CaptionText 'SIMATIC'
      DiagonalMovement <- "D_Pct"
   TextField "Label_M_D" at 814,388 size 198x16; Text 'M_D'
   Gauge "M_Direct" at 6,408 size 150x150; CaptionText 'SIMATIC'
      DirectMovement <- "D_X"
      DirectMovement <- "D_Y"
   TextField "Label_M_Direct" at 6,590 size 198x16; Text 'M_Direct'
   Gauge "E_Range" at 208,408 size 150x150; CaptionText 'SIMATIC'
      ObjectEnable <- "D_Range"
   TextField "Label_E_Range" at 208,590 size 198x16; Text 'E_Range'
   Gauge "E_Bit" at 410,408 size 150x150; CaptionText 'SIMATIC'
      ObjectEnable <- "D_En"
   TextField "Label_E_Bit" at 410,590 size 198x16; Text 'E_Bit'
   Gauge "PV_Pct" at 612,408 size 150x150; CaptionText 'SIMATIC'
      ProcessValue <- "D_Pct"
   TextField "Label_PV_Pct" at 612,590 size 198x16; Text 'PV_Pct'
   Gauge "PV_Real" at 814,408 size 150x150; CaptionText 'SIMATIC'
      ProcessValue <- "D_Real"
   TextField "Label_PV_Real" at 814,590 size 198x16; Text 'PV_Real'
   IOField "State" at 4,742 size 60x22; FormatPattern 9
      ProcessValue <- "D_State"
   Button "S1" at 70,742 size 40x22; TextOff 'S1'
      on Click: "SetS1"()
   Button "S2" at 114,742 size 40x22; TextOff 'S2'
      on Click: "SetS2"()
   Button "S3" at 158,742 size 40x22; TextOff 'S3'
      on Click: "SetS3"()
   Button "S4" at 202,742 size 40x22; TextOff 'S4'
      on Click: "SetS4"()
   Button "Next" at 980,742 size 40x22; TextOff 'Next'
      on Click: ActivateScreen("D_Gauge_2", 0)

screen "D_Gauge_2" 1024x768
   Gauge "PV_Pct_MaxMin" at 6,4 size 150x150; CaptionText 'SIMATIC'
      ProcessValue <- "D_Pct"
      MaximumValue <- "D_Max"
      MinimumValue <- "D_Min"
   TextField "Label_PV_Pct_MaxMin" at 6,186 size 198x16; Text 'PV_Pct_MaxMin'
   IOField "State" at 4,742 size 60x22; FormatPattern 9
      ProcessValue <- "D_State"
   Button "S1" at 70,742 size 40x22; TextOff 'S1'
      on Click: "SetS1"()
   Button "S2" at 114,742 size 40x22; TextOff 'S2'
      on Click: "SetS2"()
   Button "S3" at 158,742 size 40x22; TextOff 'S3'
      on Click: "SetS3"()
   Button "S4" at 202,742 size 40x22; TextOff 'S4'
      on Click: "SetS4"()
   Button "Next" at 980,742 size 40x22; TextOff 'Next'
      on Click: ActivateScreen("D_Clock_1", 0)

screen "D_GraphicIOField_1" 1024x768
   GraphicIOField "Static" at 6,4 size 60x60
   TextField "Label_Static" at 6,96 size 108x16; Text 'Static'
   GraphicIOField "A_Range" at 118,4 size 60x60
      Appearance <- "D_Range"
   TextField "Label_A_Range" at 118,96 size 108x16; Text 'A_Range'
   GraphicIOField "A_Flash" at 230,4 size 60x60
      Appearance <- "D_Range"
   TextField "Label_A_Flash" at 230,96 size 108x16; Text 'A_Flash'
   GraphicIOField "A_Bit" at 342,4 size 60x60
      Appearance <- "D_Bool"
   TextField "Label_A_Bit" at 342,96 size 108x16; Text 'A_Bit'
   GraphicIOField "A_Bits" at 454,4 size 60x60
      Appearance <- "D_Bits"
   TextField "Label_A_Bits" at 454,96 size 108x16; Text 'A_Bits'
   GraphicIOField "V_Range" at 566,4 size 60x60
      Visibility <- "D_Range"
   TextField "Label_V_Range" at 566,96 size 108x16; Text 'V_Range'
   GraphicIOField "V_Bit" at 678,4 size 60x60
      Visibility <- "D_Vis"
   TextField "Label_V_Bit" at 678,96 size 108x16; Text 'V_Bit'
   GraphicIOField "M_H" at 790,4 size 60x60
      HorizontalMovement <- "D_Pct"
   TextField "Label_M_H" at 790,96 size 108x16; Text 'M_H'
   GraphicIOField "M_V" at 902,4 size 60x60
      VerticalMovement <- "D_Pct"
   TextField "Label_M_V" at 902,96 size 108x16; Text 'M_V'
   GraphicIOField "M_D" at 6,116 size 60x60
      DiagonalMovement <- "D_Pct"
   TextField "Label_M_D" at 6,208 size 108x16; Text 'M_D'
   GraphicIOField "M_Direct" at 118,116 size 60x60
      DirectMovement <- "D_X"
      DirectMovement <- "D_Y"
   TextField "Label_M_Direct" at 118,208 size 108x16; Text 'M_Direct'
   GraphicIOField "E_Range" at 230,116 size 60x60
      ObjectEnable <- "D_Range"
   TextField "Label_E_Range" at 230,208 size 108x16; Text 'E_Range'
   GraphicIOField "E_Bit" at 342,116 size 60x60
      ObjectEnable <- "D_En"
   TextField "Label_E_Bit" at 342,208 size 108x16; Text 'E_Bit'
   IOField "State" at 4,742 size 60x22; FormatPattern 9
      ProcessValue <- "D_State"
   Button "S1" at 70,742 size 40x22; TextOff 'S1'
      on Click: "SetS1"()
   Button "S2" at 114,742 size 40x22; TextOff 'S2'
      on Click: "SetS2"()
   Button "S3" at 158,742 size 40x22; TextOff 'S3'
      on Click: "SetS3"()
   Button "S4" at 202,742 size 40x22; TextOff 'S4'
      on Click: "SetS4"()
   Button "Next" at 980,742 size 40x22; TextOff 'Next'
      on Click: ActivateScreen("D_DateTimeField_1", 0)

screen "D_GraphicView_1" 1024x768
   GraphicView "Static" at 6,4 size 100x60
   TextField "Label_Static" at 6,96 size 148x16; Text 'Static'
   GraphicView "A_Range" at 158,4 size 100x60
      Appearance <- "D_Range"
   TextField "Label_A_Range" at 158,96 size 148x16; Text 'A_Range'
   GraphicView "A_Flash" at 310,4 size 100x60
      Appearance <- "D_Range"
   TextField "Label_A_Flash" at 310,96 size 148x16; Text 'A_Flash'
   GraphicView "A_Bit" at 462,4 size 100x60
      Appearance <- "D_Bool"
   TextField "Label_A_Bit" at 462,96 size 148x16; Text 'A_Bit'
   GraphicView "A_Bits" at 614,4 size 100x60
      Appearance <- "D_Bits"
   TextField "Label_A_Bits" at 614,96 size 148x16; Text 'A_Bits'
   GraphicView "V_Range" at 766,4 size 100x60
      Visibility <- "D_Range"
   TextField "Label_V_Range" at 766,96 size 148x16; Text 'V_Range'
   GraphicView "V_Bit" at 6,116 size 100x60
      Visibility <- "D_Vis"
   TextField "Label_V_Bit" at 6,208 size 148x16; Text 'V_Bit'
   GraphicView "M_H" at 158,116 size 100x60
      HorizontalMovement <- "D_Pct"
   TextField "Label_M_H" at 158,208 size 148x16; Text 'M_H'
   GraphicView "M_V" at 310,116 size 100x60
      VerticalMovement <- "D_Pct"
   TextField "Label_M_V" at 310,208 size 148x16; Text 'M_V'
   GraphicView "M_D" at 462,116 size 100x60
      DiagonalMovement <- "D_Pct"
   TextField "Label_M_D" at 462,208 size 148x16; Text 'M_D'
   GraphicView "M_Direct" at 614,116 size 100x60
      DirectMovement <- "D_X"
      DirectMovement <- "D_Y"
   TextField "Label_M_Direct" at 614,208 size 148x16; Text 'M_Direct'
   GraphicView "E_Range" at 766,116 size 100x60
      ObjectEnable <- "D_Range"
   TextField "Label_E_Range" at 766,208 size 148x16; Text 'E_Range'
   GraphicView "E_Bit" at 6,228 size 100x60
      ObjectEnable <- "D_En"
   TextField "Label_E_Bit" at 6,320 size 148x16; Text 'E_Bit'
   IOField "State" at 4,742 size 60x22; FormatPattern 9
      ProcessValue <- "D_State"
   Button "S1" at 70,742 size 40x22; TextOff 'S1'
      on Click: "SetS1"()
   Button "S2" at 114,742 size 40x22; TextOff 'S2'
      on Click: "SetS2"()
   Button "S3" at 158,742 size 40x22; TextOff 'S3'
      on Click: "SetS3"()
   Button "S4" at 202,742 size 40x22; TextOff 'S4'
      on Click: "SetS4"()
   Button "Next" at 980,742 size 40x22; TextOff 'Next'
      on Click: ActivateScreen("D_IOField_1", 0)

screen "D_IOField_1" 1024x768
   IOField "Static" at 6,4 size 100x30
   TextField "Label_Static" at 6,66 size 148x16; Text 'Static'
   IOField "A_Range" at 158,4 size 100x30
      Appearance <- "D_Range"
   TextField "Label_A_Range" at 158,66 size 148x16; Text 'A_Range'
   IOField "A_Flash" at 310,4 size 100x30
      Appearance <- "D_Range"
   TextField "Label_A_Flash" at 310,66 size 148x16; Text 'A_Flash'
   IOField "A_Bit" at 462,4 size 100x30
      Appearance <- "D_Bool"
   TextField "Label_A_Bit" at 462,66 size 148x16; Text 'A_Bit'
   IOField "A_Bits" at 614,4 size 100x30
      Appearance <- "D_Bits"
   TextField "Label_A_Bits" at 614,66 size 148x16; Text 'A_Bits'
   IOField "V_Range" at 766,4 size 100x30
      Visibility <- "D_Range"
   TextField "Label_V_Range" at 766,66 size 148x16; Text 'V_Range'
   IOField "V_Bit" at 6,86 size 100x30
      Visibility <- "D_Vis"
   TextField "Label_V_Bit" at 6,148 size 148x16; Text 'V_Bit'
   IOField "M_H" at 158,86 size 100x30
      HorizontalMovement <- "D_Pct"
   TextField "Label_M_H" at 158,148 size 148x16; Text 'M_H'
   IOField "M_V" at 310,86 size 100x30
      VerticalMovement <- "D_Pct"
   TextField "Label_M_V" at 310,148 size 148x16; Text 'M_V'
   IOField "M_D" at 462,86 size 100x30
      DiagonalMovement <- "D_Pct"
   TextField "Label_M_D" at 462,148 size 148x16; Text 'M_D'
   IOField "M_Direct" at 614,86 size 100x30
      DirectMovement <- "D_X"
      DirectMovement <- "D_Y"
   TextField "Label_M_Direct" at 614,148 size 148x16; Text 'M_Direct'
   IOField "E_Range" at 766,86 size 100x30
      ObjectEnable <- "D_Range"
   TextField "Label_E_Range" at 766,148 size 148x16; Text 'E_Range'
   IOField "E_Bit" at 6,168 size 100x30
      ObjectEnable <- "D_En"
   TextField "Label_E_Bit" at 6,230 size 148x16; Text 'E_Bit'
   IOField "PV_SInt" at 158,168 size 100x30; FormatPattern s999
      ProcessValue <- "D_SInt"
   TextField "Label_PV_SInt" at 158,230 size 148x16; Text 'PV_SInt'
   IOField "PV_Int" at 310,168 size 100x30; FormatPattern s99999
      ProcessValue <- "D_Int"
   TextField "Label_PV_Int" at 310,230 size 148x16; Text 'PV_Int'
   IOField "PV_DInt" at 462,168 size 100x30; FormatPattern s9999999999
      ProcessValue <- "D_DInt"
   TextField "Label_PV_DInt" at 462,230 size 148x16; Text 'PV_DInt'
   IOField "PV_USInt" at 614,168 size 100x30; FormatPattern 999
      ProcessValue <- "D_USInt"
   TextField "Label_PV_USInt" at 614,230 size 148x16; Text 'PV_USInt'
   IOField "PV_UInt" at 766,168 size 100x30; FormatPattern 99999
      ProcessValue <- "D_UInt"
   TextField "Label_PV_UInt" at 766,230 size 148x16; Text 'PV_UInt'
   IOField "PV_UDInt" at 6,250 size 100x30; FormatPattern 9999999999
      ProcessValue <- "D_UDInt"
   TextField "Label_PV_UDInt" at 6,312 size 148x16; Text 'PV_UDInt'
   IOField "PV_Real" at 158,250 size 100x30
      ProcessValue <- "D_Real"
   TextField "Label_PV_Real" at 158,312 size 148x16; Text 'PV_Real'
   IOField "PV_LReal" at 310,250 size 100x30
      ProcessValue <- "D_LReal"
   TextField "Label_PV_LReal" at 310,312 size 148x16; Text 'PV_LReal'
   IOField "PV_String" at 462,250 size 100x30
      ProcessValue <- "D_String"
   TextField "Label_PV_String" at 462,312 size 148x16; Text 'PV_String'
   IOField "PV_Int_Shift2" at 614,250 size 100x30; FormatPattern s99999
      ProcessValue <- "D_Int"
   TextField "Label_PV_Int_Shift2" at 614,312 size 148x16; Text 'PV_Int_Shift2'
   IOField "PV_Int_s999999" at 766,250 size 100x30; FormatPattern s999999
      ProcessValue <- "D_Int"
   TextField "Label_PV_Int_s999999" at 766,312 size 148x16; Text 'PV_Int_s999999'
   IOField "PV_Real_s9999_99" at 6,332 size 100x30; FormatPattern s9999.99
      ProcessValue <- "D_Real"
   TextField "Label_PV_Real_s9999_99" at 6,394 size 148x16; Text 'PV_Real_s9999_99'
   IOField "PV_Int_Output" at 158,332 size 100x30; FormatPattern s99999
      ProcessValue <- "D_Int"
   TextField "Label_PV_Int_Output" at 158,394 size 148x16; Text 'PV_Int_Output'
   IOField "PV_Int_s99" at 310,332 size 100x30; FormatPattern s99
      ProcessValue <- "D_Int"
   TextField "Label_PV_Int_s99" at 310,394 size 148x16; Text 'PV_Int_s99'
   IOField "State" at 4,742 size 60x22; FormatPattern 9
      ProcessValue <- "D_State"
   Button "S1" at 70,742 size 40x22; TextOff 'S1'
      on Click: "SetS1"()
   Button "S2" at 114,742 size 40x22; TextOff 'S2'
      on Click: "SetS2"()
   Button "S3" at 158,742 size 40x22; TextOff 'S3'
      on Click: "SetS3"()
   Button "S4" at 202,742 size 40x22; TextOff 'S4'
      on Click: "SetS4"()
   Button "Next" at 980,742 size 40x22; TextOff 'Next'
      on Click: ActivateScreen("D_Button_1", 0)

screen "D_Line_1" 1024x768
   TextField "Label_Static" at 6,86 size 148x16; Text 'Static'
   Line "A_Range" at 158,4 size 100x50
      Appearance <- "D_Range"
   TextField "Label_A_Range" at 158,86 size 148x16; Text 'A_Range'
   Line "A_Flash" at 310,4 size 100x50
      Appearance <- "D_Range"
   TextField "Label_A_Flash" at 310,86 size 148x16; Text 'A_Flash'
   Line "A_Bit" at 462,4 size 100x50
      Appearance <- "D_Bool"
   TextField "Label_A_Bit" at 462,86 size 148x16; Text 'A_Bit'
   Line "A_Bits" at 614,4 size 100x50
      Appearance <- "D_Bits"
   TextField "Label_A_Bits" at 614,86 size 148x16; Text 'A_Bits'
   Line "V_Range" at 766,4 size 100x50
      Visibility <- "D_Range"
   TextField "Label_V_Range" at 766,86 size 148x16; Text 'V_Range'
   Line "V_Bit" at 6,106 size 100x50
      Visibility <- "D_Vis"
   TextField "Label_V_Bit" at 6,188 size 148x16; Text 'V_Bit'
   Line "M_H" at 158,106 size 100x50
      HorizontalMovement <- "D_Pct"
   TextField "Label_M_H" at 158,188 size 148x16; Text 'M_H'
   Line "M_V" at 310,106 size 100x50
      VerticalMovement <- "D_Pct"
   TextField "Label_M_V" at 310,188 size 148x16; Text 'M_V'
   Line "M_D" at 462,106 size 100x50
      DiagonalMovement <- "D_Pct"
   TextField "Label_M_D" at 462,188 size 148x16; Text 'M_D'
   Line "M_Direct" at 614,106 size 100x50
      DirectMovement <- "D_X"
      DirectMovement <- "D_Y"
   TextField "Label_M_Direct" at 614,188 size 148x16; Text 'M_Direct'
   Line "E_Range" at 766,106 size 100x50
      ObjectEnable <- "D_Range"
   TextField "Label_E_Range" at 766,188 size 148x16; Text 'E_Range'
   Line "E_Bit" at 6,208 size 100x50
      ObjectEnable <- "D_En"
   TextField "Label_E_Bit" at 6,290 size 148x16; Text 'E_Bit'
   IOField "State" at 4,742 size 60x22; FormatPattern 9
      ProcessValue <- "D_State"
   Button "S1" at 70,742 size 40x22; TextOff 'S1'
      on Click: "SetS1"()
   Button "S2" at 114,742 size 40x22; TextOff 'S2'
      on Click: "SetS2"()
   Button "S3" at 158,742 size 40x22; TextOff 'S3'
      on Click: "SetS3"()
   Button "S4" at 202,742 size 40x22; TextOff 'S4'
      on Click: "SetS4"()
   Button "Next" at 980,742 size 40x22; TextOff 'Next'
      on Click: ActivateScreen("D_Polyline_1", 0)

screen "D_Polygon_1" 1024x768
   TextField "Label_Static" at 6,86 size 148x16; Text 'Static'
   Polygon "A_Range" at 158,4 size 100x50
      Appearance <- "D_Range"
   TextField "Label_A_Range" at 158,86 size 148x16; Text 'A_Range'
   Polygon "A_Flash" at 310,4 size 100x50
      Appearance <- "D_Range"
   TextField "Label_A_Flash" at 310,86 size 148x16; Text 'A_Flash'
   Polygon "A_Bit" at 462,4 size 100x50
      Appearance <- "D_Bool"
   TextField "Label_A_Bit" at 462,86 size 148x16; Text 'A_Bit'
   Polygon "A_Bits" at 614,4 size 100x50
      Appearance <- "D_Bits"
   TextField "Label_A_Bits" at 614,86 size 148x16; Text 'A_Bits'
   Polygon "V_Range" at 766,4 size 100x50
      Visibility <- "D_Range"
   TextField "Label_V_Range" at 766,86 size 148x16; Text 'V_Range'
   Polygon "V_Bit" at 6,106 size 100x50
      Visibility <- "D_Vis"
   TextField "Label_V_Bit" at 6,188 size 148x16; Text 'V_Bit'
   Polygon "M_H" at 158,106 size 100x50
      HorizontalMovement <- "D_Pct"
   TextField "Label_M_H" at 158,188 size 148x16; Text 'M_H'
   Polygon "M_V" at 310,106 size 100x50
      VerticalMovement <- "D_Pct"
   TextField "Label_M_V" at 310,188 size 148x16; Text 'M_V'
   Polygon "M_D" at 462,106 size 100x50
      DiagonalMovement <- "D_Pct"
   TextField "Label_M_D" at 462,188 size 148x16; Text 'M_D'
   Polygon "M_Direct" at 614,106 size 100x50
      DirectMovement <- "D_X"
      DirectMovement <- "D_Y"
   TextField "Label_M_Direct" at 614,188 size 148x16; Text 'M_Direct'
   Polygon "E_Range" at 766,106 size 100x50
      ObjectEnable <- "D_Range"
   TextField "Label_E_Range" at 766,188 size 148x16; Text 'E_Range'
   Polygon "E_Bit" at 6,208 size 100x50
      ObjectEnable <- "D_En"
   TextField "Label_E_Bit" at 6,290 size 148x16; Text 'E_Bit'
   IOField "State" at 4,742 size 60x22; FormatPattern 9
      ProcessValue <- "D_State"
   Button "S1" at 70,742 size 40x22; TextOff 'S1'
      on Click: "SetS1"()
   Button "S2" at 114,742 size 40x22; TextOff 'S2'
      on Click: "SetS2"()
   Button "S3" at 158,742 size 40x22; TextOff 'S3'
      on Click: "SetS3"()
   Button "S4" at 202,742 size 40x22; TextOff 'S4'
      on Click: "SetS4"()
   Button "Next" at 980,742 size 40x22; TextOff 'Next'
      on Click: ActivateScreen("D_Ellipse_1", 0)

screen "D_Polyline_1" 1024x768
   TextField "Label_Static" at 6,86 size 148x16; Text 'Static'
   Polyline "A_Range" at 158,4 size 100x50
      Appearance <- "D_Range"
   TextField "Label_A_Range" at 158,86 size 148x16; Text 'A_Range'
   Polyline "A_Flash" at 310,4 size 100x50
      Appearance <- "D_Range"
   TextField "Label_A_Flash" at 310,86 size 148x16; Text 'A_Flash'
   Polyline "A_Bit" at 462,4 size 100x50
      Appearance <- "D_Bool"
   TextField "Label_A_Bit" at 462,86 size 148x16; Text 'A_Bit'
   Polyline "A_Bits" at 614,4 size 100x50
      Appearance <- "D_Bits"
   TextField "Label_A_Bits" at 614,86 size 148x16; Text 'A_Bits'
   Polyline "V_Range" at 766,4 size 100x50
      Visibility <- "D_Range"
   TextField "Label_V_Range" at 766,86 size 148x16; Text 'V_Range'
   Polyline "V_Bit" at 6,106 size 100x50
      Visibility <- "D_Vis"
   TextField "Label_V_Bit" at 6,188 size 148x16; Text 'V_Bit'
   Polyline "M_H" at 158,106 size 100x50
      HorizontalMovement <- "D_Pct"
   TextField "Label_M_H" at 158,188 size 148x16; Text 'M_H'
   Polyline "M_V" at 310,106 size 100x50
      VerticalMovement <- "D_Pct"
   TextField "Label_M_V" at 310,188 size 148x16; Text 'M_V'
   Polyline "M_D" at 462,106 size 100x50
      DiagonalMovement <- "D_Pct"
   TextField "Label_M_D" at 462,188 size 148x16; Text 'M_D'
   Polyline "M_Direct" at 614,106 size 100x50
      DirectMovement <- "D_X"
      DirectMovement <- "D_Y"
   TextField "Label_M_Direct" at 614,188 size 148x16; Text 'M_Direct'
   Polyline "E_Range" at 766,106 size 100x50
      ObjectEnable <- "D_Range"
   TextField "Label_E_Range" at 766,188 size 148x16; Text 'E_Range'
   Polyline "E_Bit" at 6,208 size 100x50
      ObjectEnable <- "D_En"
   TextField "Label_E_Bit" at 6,290 size 148x16; Text 'E_Bit'
   IOField "State" at 4,742 size 60x22; FormatPattern 9
      ProcessValue <- "D_State"
   Button "S1" at 70,742 size 40x22; TextOff 'S1'
      on Click: "SetS1"()
   Button "S2" at 114,742 size 40x22; TextOff 'S2'
      on Click: "SetS2"()
   Button "S3" at 158,742 size 40x22; TextOff 'S3'
      on Click: "SetS3"()
   Button "S4" at 202,742 size 40x22; TextOff 'S4'
      on Click: "SetS4"()
   Button "Next" at 980,742 size 40x22; TextOff 'Next'
      on Click: ActivateScreen("D_Polygon_1", 0)

screen "D_Rectangle_1" 1024x768
   TextField "Label_Static" at 6,86 size 148x16; Text 'Static'
   Rectangle "A_Range" at 158,4 size 100x50
      Appearance <- "D_Range"
   TextField "Label_A_Range" at 158,86 size 148x16; Text 'A_Range'
   Rectangle "A_Flash" at 310,4 size 100x50
      Appearance <- "D_Range"
   TextField "Label_A_Flash" at 310,86 size 148x16; Text 'A_Flash'
   Rectangle "A_Bit" at 462,4 size 100x50
      Appearance <- "D_Bool"
   TextField "Label_A_Bit" at 462,86 size 148x16; Text 'A_Bit'
   Rectangle "A_Bits" at 614,4 size 100x50
      Appearance <- "D_Bits"
   TextField "Label_A_Bits" at 614,86 size 148x16; Text 'A_Bits'
   Rectangle "V_Range" at 766,4 size 100x50
      Visibility <- "D_Range"
   TextField "Label_V_Range" at 766,86 size 148x16; Text 'V_Range'
   Rectangle "V_Bit" at 6,106 size 100x50
      Visibility <- "D_Vis"
   TextField "Label_V_Bit" at 6,188 size 148x16; Text 'V_Bit'
   Rectangle "M_H" at 158,106 size 100x50
      HorizontalMovement <- "D_Pct"
   TextField "Label_M_H" at 158,188 size 148x16; Text 'M_H'
   Rectangle "M_V" at 310,106 size 100x50
      VerticalMovement <- "D_Pct"
   TextField "Label_M_V" at 310,188 size 148x16; Text 'M_V'
   Rectangle "M_D" at 462,106 size 100x50
      DiagonalMovement <- "D_Pct"
   TextField "Label_M_D" at 462,188 size 148x16; Text 'M_D'
   Rectangle "M_Direct" at 614,106 size 100x50
      DirectMovement <- "D_X"
      DirectMovement <- "D_Y"
   TextField "Label_M_Direct" at 614,188 size 148x16; Text 'M_Direct'
   Rectangle "E_Range" at 766,106 size 100x50
      ObjectEnable <- "D_Range"
   TextField "Label_E_Range" at 766,188 size 148x16; Text 'E_Range'
   Rectangle "E_Bit" at 6,208 size 100x50
      ObjectEnable <- "D_En"
   TextField "Label_E_Bit" at 6,290 size 148x16; Text 'E_Bit'
   IOField "State" at 4,742 size 60x22; FormatPattern 9
      ProcessValue <- "D_State"
   Button "S1" at 70,742 size 40x22; TextOff 'S1'
      on Click: "SetS1"()
   Button "S2" at 114,742 size 40x22; TextOff 'S2'
      on Click: "SetS2"()
   Button "S3" at 158,742 size 40x22; TextOff 'S3'
      on Click: "SetS3"()
   Button "S4" at 202,742 size 40x22; TextOff 'S4'
      on Click: "SetS4"()
   Button "Next" at 980,742 size 40x22; TextOff 'Next'
      on Click: ActivateScreen("D_TextField_1", 0)

screen "D_Slider_1" 1024x768
   Slider "Static" at 6,4 size 60x160; Caption 'SIMATIC'
   TextField "Label_Static" at 6,196 size 108x16; Text 'Static'
   Slider "A_Range" at 118,4 size 60x160; Caption 'SIMATIC'
      Appearance <- "D_Range"
   TextField "Label_A_Range" at 118,196 size 108x16; Text 'A_Range'
   Slider "A_Flash" at 230,4 size 60x160; Caption 'SIMATIC'
      Appearance <- "D_Range"
   TextField "Label_A_Flash" at 230,196 size 108x16; Text 'A_Flash'
   Slider "A_Bit" at 342,4 size 60x160; Caption 'SIMATIC'
      Appearance <- "D_Bool"
   TextField "Label_A_Bit" at 342,196 size 108x16; Text 'A_Bit'
   Slider "A_Bits" at 454,4 size 60x160; Caption 'SIMATIC'
      Appearance <- "D_Bits"
   TextField "Label_A_Bits" at 454,196 size 108x16; Text 'A_Bits'
   Slider "V_Range" at 566,4 size 60x160; Caption 'SIMATIC'
      Visibility <- "D_Range"
   TextField "Label_V_Range" at 566,196 size 108x16; Text 'V_Range'
   Slider "V_Bit" at 678,4 size 60x160; Caption 'SIMATIC'
      Visibility <- "D_Vis"
   TextField "Label_V_Bit" at 678,196 size 108x16; Text 'V_Bit'
   Slider "M_H" at 790,4 size 60x160; Caption 'SIMATIC'
      HorizontalMovement <- "D_Pct"
   TextField "Label_M_H" at 790,196 size 108x16; Text 'M_H'
   Slider "M_V" at 902,4 size 60x160; Caption 'SIMATIC'
      VerticalMovement <- "D_Pct"
   TextField "Label_M_V" at 902,196 size 108x16; Text 'M_V'
   Slider "M_D" at 6,216 size 60x160; Caption 'SIMATIC'
      DiagonalMovement <- "D_Pct"
   TextField "Label_M_D" at 6,408 size 108x16; Text 'M_D'
   Slider "M_Direct" at 118,216 size 60x160; Caption 'SIMATIC'
      DirectMovement <- "D_X"
      DirectMovement <- "D_Y"
   TextField "Label_M_Direct" at 118,408 size 108x16; Text 'M_Direct'
   Slider "E_Range" at 230,216 size 60x160; Caption 'SIMATIC'
      ObjectEnable <- "D_Range"
   TextField "Label_E_Range" at 230,408 size 108x16; Text 'E_Range'
   Slider "E_Bit" at 342,216 size 60x160; Caption 'SIMATIC'
      ObjectEnable <- "D_En"
   TextField "Label_E_Bit" at 342,408 size 108x16; Text 'E_Bit'
   Slider "PV_Pct" at 454,216 size 60x160; Caption 'SIMATIC'
      ProcessValue <- "D_Pct"
   TextField "Label_PV_Pct" at 454,408 size 108x16; Text 'PV_Pct'
   Slider "PV_Int" at 566,216 size 60x160; Caption 'SIMATIC'
      ProcessValue <- "D_Int"
   TextField "Label_PV_Int" at 566,408 size 108x16; Text 'PV_Int'
   Slider "PV_Pct_0_200" at 678,216 size 60x160; Caption 'SIMATIC'
      ProcessValue <- "D_Pct"
   TextField "Label_PV_Pct_0_200" at 678,408 size 108x16; Text 'PV_Pct_0_200'
   IOField "State" at 4,742 size 60x22; FormatPattern 9
      ProcessValue <- "D_State"
   Button "S1" at 70,742 size 40x22; TextOff 'S1'
      on Click: "SetS1"()
   Button "S2" at 114,742 size 40x22; TextOff 'S2'
      on Click: "SetS2"()
   Button "S3" at 158,742 size 40x22; TextOff 'S3'
      on Click: "SetS3"()
   Button "S4" at 202,742 size 40x22; TextOff 'S4'
      on Click: "SetS4"()
   Button "Next" at 980,742 size 40x22; TextOff 'Next'
      on Click: ActivateScreen("D_Gauge_1", 0)

screen "D_Switch_1" 1024x768
   Switch "Static" at 6,4 size 120x40; CaptionText 'Switch'; TextOff '0'; TextOn '1'
   TextField "Label_Static" at 6,76 size 168x16; Text 'Static'
   Switch "A_Range" at 178,4 size 120x40; CaptionText 'Switch'; TextOff '0'; TextOn '1'
      Appearance <- "D_Range"
   TextField "Label_A_Range" at 178,76 size 168x16; Text 'A_Range'
   Switch "A_Flash" at 350,4 size 120x40; CaptionText 'Switch'; TextOff '0'; TextOn '1'
      Appearance <- "D_Range"
   TextField "Label_A_Flash" at 350,76 size 168x16; Text 'A_Flash'
   Switch "A_Bit" at 522,4 size 120x40; CaptionText 'Switch'; TextOff '0'; TextOn '1'
      Appearance <- "D_Bool"
   TextField "Label_A_Bit" at 522,76 size 168x16; Text 'A_Bit'
   Switch "A_Bits" at 694,4 size 120x40; CaptionText 'Switch'; TextOff '0'; TextOn '1'
      Appearance <- "D_Bits"
   TextField "Label_A_Bits" at 694,76 size 168x16; Text 'A_Bits'
   Switch "V_Range" at 6,96 size 120x40; CaptionText 'Switch'; TextOff '0'; TextOn '1'
      Visibility <- "D_Range"
   TextField "Label_V_Range" at 6,168 size 168x16; Text 'V_Range'
   Switch "V_Bit" at 178,96 size 120x40; CaptionText 'Switch'; TextOff '0'; TextOn '1'
      Visibility <- "D_Vis"
   TextField "Label_V_Bit" at 178,168 size 168x16; Text 'V_Bit'
   Switch "M_H" at 350,96 size 120x40; CaptionText 'Switch'; TextOff '0'; TextOn '1'
      HorizontalMovement <- "D_Pct"
   TextField "Label_M_H" at 350,168 size 168x16; Text 'M_H'
   Switch "M_V" at 522,96 size 120x40; CaptionText 'Switch'; TextOff '0'; TextOn '1'
      VerticalMovement <- "D_Pct"
   TextField "Label_M_V" at 522,168 size 168x16; Text 'M_V'
   Switch "M_D" at 694,96 size 120x40; CaptionText 'Switch'; TextOff '0'; TextOn '1'
      DiagonalMovement <- "D_Pct"
   TextField "Label_M_D" at 694,168 size 168x16; Text 'M_D'
   Switch "M_Direct" at 6,188 size 120x40; CaptionText 'Switch'; TextOff '0'; TextOn '1'
      DirectMovement <- "D_X"
      DirectMovement <- "D_Y"
   TextField "Label_M_Direct" at 6,260 size 168x16; Text 'M_Direct'
   Switch "E_Range" at 178,188 size 120x40; CaptionText 'Switch'; TextOff '0'; TextOn '1'
      ObjectEnable <- "D_Range"
   TextField "Label_E_Range" at 178,260 size 168x16; Text 'E_Range'
   Switch "E_Bit" at 350,188 size 120x40; CaptionText 'Switch'; TextOff '0'; TextOn '1'
      ObjectEnable <- "D_En"
   TextField "Label_E_Bit" at 350,260 size 168x16; Text 'E_Bit'
   Switch "PV_Bool" at 522,188 size 120x40; CaptionText 'Switch'; TextOff '0'; TextOn '1'
      ProcessValue <- "D_Bool"
   TextField "Label_PV_Bool" at 522,260 size 168x16; Text 'PV_Bool'
   IOField "State" at 4,742 size 60x22; FormatPattern 9
      ProcessValue <- "D_State"
   Button "S1" at 70,742 size 40x22; TextOff 'S1'
      on Click: "SetS1"()
   Button "S2" at 114,742 size 40x22; TextOff 'S2'
      on Click: "SetS2"()
   Button "S3" at 158,742 size 40x22; TextOff 'S3'
      on Click: "SetS3"()
   Button "S4" at 202,742 size 40x22; TextOff 'S4'
      on Click: "SetS4"()
   Button "Next" at 980,742 size 40x22; TextOff 'Next'
      on Click: ActivateScreen("D_SymbolLibrary_1", 0)

screen "D_SymbolicIOField_1" 1024x768
   SymbolicIOField "Static" at 6,4 size 120x30; TextOff '0'; TextOn '1'
   TextField "Label_Static" at 6,66 size 168x16; Text 'Static'
   SymbolicIOField "A_Range" at 178,4 size 120x30; TextOff '0'; TextOn '1'
      Appearance <- "D_Range"
   TextField "Label_A_Range" at 178,66 size 168x16; Text 'A_Range'
   SymbolicIOField "A_Flash" at 350,4 size 120x30; TextOff '0'; TextOn '1'
      Appearance <- "D_Range"
   TextField "Label_A_Flash" at 350,66 size 168x16; Text 'A_Flash'
   SymbolicIOField "A_Bit" at 522,4 size 120x30; TextOff '0'; TextOn '1'
      Appearance <- "D_Bool"
   TextField "Label_A_Bit" at 522,66 size 168x16; Text 'A_Bit'
   SymbolicIOField "A_Bits" at 694,4 size 120x30; TextOff '0'; TextOn '1'
      Appearance <- "D_Bits"
   TextField "Label_A_Bits" at 694,66 size 168x16; Text 'A_Bits'
   SymbolicIOField "V_Range" at 6,86 size 120x30; TextOff '0'; TextOn '1'
      Visibility <- "D_Range"
   TextField "Label_V_Range" at 6,148 size 168x16; Text 'V_Range'
   SymbolicIOField "V_Bit" at 178,86 size 120x30; TextOff '0'; TextOn '1'
      Visibility <- "D_Vis"
   TextField "Label_V_Bit" at 178,148 size 168x16; Text 'V_Bit'
   SymbolicIOField "M_H" at 350,86 size 120x30; TextOff '0'; TextOn '1'
      HorizontalMovement <- "D_Pct"
   TextField "Label_M_H" at 350,148 size 168x16; Text 'M_H'
   SymbolicIOField "M_V" at 522,86 size 120x30; TextOff '0'; TextOn '1'
      VerticalMovement <- "D_Pct"
   TextField "Label_M_V" at 522,148 size 168x16; Text 'M_V'
   SymbolicIOField "M_D" at 694,86 size 120x30; TextOff '0'; TextOn '1'
      DiagonalMovement <- "D_Pct"
   TextField "Label_M_D" at 694,148 size 168x16; Text 'M_D'
   SymbolicIOField "M_Direct" at 6,168 size 120x30; TextOff '0'; TextOn '1'
      DirectMovement <- "D_X"
      DirectMovement <- "D_Y"
   TextField "Label_M_Direct" at 6,230 size 168x16; Text 'M_Direct'
   SymbolicIOField "E_Range" at 178,168 size 120x30; TextOff '0'; TextOn '1'
      ObjectEnable <- "D_Range"
   TextField "Label_E_Range" at 178,230 size 168x16; Text 'E_Range'
   SymbolicIOField "E_Bit" at 350,168 size 120x30; TextOff '0'; TextOn '1'
      ObjectEnable <- "D_En"
   TextField "Label_E_Bit" at 350,230 size 168x16; Text 'E_Bit'
   SymbolicIOField "PV_TL_Value" at 522,168 size 120x30; TextOff '0'; TextOn '1'; TextList "TL_Value"
      ProcessValue <- "D_TL"
   TextField "Label_PV_TL_Value" at 522,230 size 168x16; Text 'PV_TL_Value'
   SymbolicIOField "PV_TL_Bit" at 694,168 size 120x30; TextOff '0'; TextOn '1'; TextList "TL_Bit"
      ProcessValue <- "D_Bool"
   TextField "Label_PV_TL_Bit" at 694,230 size 168x16; Text 'PV_TL_Bit'
   SymbolicIOField "PV_TL_BitNo" at 6,250 size 120x30; TextOff '0'; TextOn '1'; TextList "TL_BitNo"
      ProcessValue <- "D_Bits"
   TextField "Label_PV_TL_BitNo" at 6,312 size 168x16; Text 'PV_TL_BitNo'
   IOField "State" at 4,742 size 60x22; FormatPattern 9
      ProcessValue <- "D_State"
   Button "S1" at 70,742 size 40x22; TextOff 'S1'
      on Click: "SetS1"()
   Button "S2" at 114,742 size 40x22; TextOff 'S2'
      on Click: "SetS2"()
   Button "S3" at 158,742 size 40x22; TextOff 'S3'
      on Click: "SetS3"()
   Button "S4" at 202,742 size 40x22; TextOff 'S4'
      on Click: "SetS4"()
   Button "Next" at 980,742 size 40x22; TextOff 'Next'
      on Click: ActivateScreen("D_GraphicIOField_1", 0)

screen "D_SymbolLibrary_1" 1024x768
   SymbolLibrary "Static" at 6,4 size 60x60
   TextField "Label_Static" at 6,96 size 108x16; Text 'Static'
   SymbolLibrary "A_Range" at 118,4 size 60x60
      Appearance <- "D_Range"
   TextField "Label_A_Range" at 118,96 size 108x16; Text 'A_Range'
   SymbolLibrary "A_Flash" at 230,4 size 60x60
      Appearance <- "D_Range"
   TextField "Label_A_Flash" at 230,96 size 108x16; Text 'A_Flash'
   SymbolLibrary "A_Bit" at 342,4 size 60x60
      Appearance <- "D_Bool"
   TextField "Label_A_Bit" at 342,96 size 108x16; Text 'A_Bit'
   SymbolLibrary "A_Bits" at 454,4 size 60x60
      Appearance <- "D_Bits"
   TextField "Label_A_Bits" at 454,96 size 108x16; Text 'A_Bits'
   SymbolLibrary "V_Range" at 566,4 size 60x60
      Visibility <- "D_Range"
   TextField "Label_V_Range" at 566,96 size 108x16; Text 'V_Range'
   SymbolLibrary "V_Bit" at 678,4 size 60x60
      Visibility <- "D_Vis"
   TextField "Label_V_Bit" at 678,96 size 108x16; Text 'V_Bit'
   SymbolLibrary "M_H" at 790,4 size 60x60
      HorizontalMovement <- "D_Pct"
   TextField "Label_M_H" at 790,96 size 108x16; Text 'M_H'
   SymbolLibrary "M_V" at 902,4 size 60x60
      VerticalMovement <- "D_Pct"
   TextField "Label_M_V" at 902,96 size 108x16; Text 'M_V'
   SymbolLibrary "M_D" at 6,116 size 60x60
      DiagonalMovement <- "D_Pct"
   TextField "Label_M_D" at 6,208 size 108x16; Text 'M_D'
   SymbolLibrary "M_Direct" at 118,116 size 60x60
      DirectMovement <- "D_X"
      DirectMovement <- "D_Y"
   TextField "Label_M_Direct" at 118,208 size 108x16; Text 'M_Direct'
   SymbolLibrary "E_Range" at 230,116 size 60x60
      ObjectEnable <- "D_Range"
   TextField "Label_E_Range" at 230,208 size 108x16; Text 'E_Range'
   SymbolLibrary "E_Bit" at 342,116 size 60x60
      ObjectEnable <- "D_En"
   TextField "Label_E_Bit" at 342,208 size 108x16; Text 'E_Bit'
   SymbolLibrary "PV_Pct" at 454,116 size 60x60
      ProcessValue <- "D_Pct"
   TextField "Label_PV_Pct" at 454,208 size 108x16; Text 'PV_Pct'
   IOField "State" at 4,742 size 60x22; FormatPattern 9
      ProcessValue <- "D_State"
   Button "S1" at 70,742 size 40x22; TextOff 'S1'
      on Click: "SetS1"()
   Button "S2" at 114,742 size 40x22; TextOff 'S2'
      on Click: "SetS2"()
   Button "S3" at 158,742 size 40x22; TextOff 'S3'
      on Click: "SetS3"()
   Button "S4" at 202,742 size 40x22; TextOff 'S4'
      on Click: "SetS4"()
   Button "Next" at 980,742 size 40x22; TextOff 'Next'
      on Click: ActivateScreen("D_Slider_1", 0)

screen "D_TextField_1" 1024x768
   TextField "Static" at 6,4 size 100x30; Text 'Text'
   TextField "Label_Static" at 6,66 size 148x16; Text 'Static'
   TextField "A_Range" at 158,4 size 100x30; Text 'Text'
      Appearance <- "D_Range"
   TextField "Label_A_Range" at 158,66 size 148x16; Text 'A_Range'
   TextField "A_Flash" at 310,4 size 100x30; Text 'Text'
      Appearance <- "D_Range"
   TextField "Label_A_Flash" at 310,66 size 148x16; Text 'A_Flash'
   TextField "A_Bit" at 462,4 size 100x30; Text 'Text'
      Appearance <- "D_Bool"
   TextField "Label_A_Bit" at 462,66 size 148x16; Text 'A_Bit'
   TextField "A_Bits" at 614,4 size 100x30; Text 'Text'
      Appearance <- "D_Bits"
   TextField "Label_A_Bits" at 614,66 size 148x16; Text 'A_Bits'
   TextField "V_Range" at 766,4 size 100x30; Text 'Text'
      Visibility <- "D_Range"
   TextField "Label_V_Range" at 766,66 size 148x16; Text 'V_Range'
   TextField "V_Bit" at 6,86 size 100x30; Text 'Text'
      Visibility <- "D_Vis"
   TextField "Label_V_Bit" at 6,148 size 148x16; Text 'V_Bit'
   TextField "M_H" at 158,86 size 100x30; Text 'Text'
      HorizontalMovement <- "D_Pct"
   TextField "Label_M_H" at 158,148 size 148x16; Text 'M_H'
   TextField "M_V" at 310,86 size 100x30; Text 'Text'
      VerticalMovement <- "D_Pct"
   TextField "Label_M_V" at 310,148 size 148x16; Text 'M_V'
   TextField "M_D" at 462,86 size 100x30; Text 'Text'
      DiagonalMovement <- "D_Pct"
   TextField "Label_M_D" at 462,148 size 148x16; Text 'M_D'
   TextField "M_Direct" at 614,86 size 100x30; Text 'Text'
      DirectMovement <- "D_X"
      DirectMovement <- "D_Y"
   TextField "Label_M_Direct" at 614,148 size 148x16; Text 'M_Direct'
   TextField "E_Range" at 766,86 size 100x30; Text 'Text'
      ObjectEnable <- "D_Range"
   TextField "Label_E_Range" at 766,148 size 148x16; Text 'E_Range'
   TextField "E_Bit" at 6,168 size 100x30; Text 'Text'
      ObjectEnable <- "D_En"
   TextField "Label_E_Bit" at 6,230 size 148x16; Text 'E_Bit'
   IOField "State" at 4,742 size 60x22; FormatPattern 9
      ProcessValue <- "D_State"
   Button "S1" at 70,742 size 40x22; TextOff 'S1'
      on Click: "SetS1"()
   Button "S2" at 114,742 size 40x22; TextOff 'S2'
      on Click: "SetS2"()
   Button "S3" at 158,742 size 40x22; TextOff 'S3'
      on Click: "SetS3"()
   Button "S4" at 202,742 size 40x22; TextOff 'S4'
      on Click: "SetS4"()
   Button "Next" at 980,742 size 40x22; TextOff 'Next'
      on Click: ActivateScreen("D_GraphicView_1", 0)

VB script "SetS1"
   SmartTags("D_State") = 1
   SmartTags("D_Bool") = False
   SmartTags("D_SInt") = -128
   SmartTags("D_Int") = -32768
   SmartTags("D_DInt") = -2147483648
   SmartTags("D_USInt") = 0
   SmartTags("D_UInt") = 0
   SmartTags("D_UDInt") = 0
   SmartTags("D_Real") = -999.999
   SmartTags("D_LReal") = -0.00000015
   SmartTags("D_String") = ""
   SmartTags("D_DateTime") = DateSerial(1990, 1, 1) + TimeSerial(0, 0, 0)
   SmartTags("D_Pct") = 0
   SmartTags("D_Range") = 5
   SmartTags("D_Bits") = 1
   SmartTags("D_Vis") = False
   SmartTags("D_En") = False
   SmartTags("D_X") = 10
   SmartTags("D_Y") = 10
   SmartTags("D_Max") = 100
   SmartTags("D_Min") = 0
   SmartTags("D_TL") = -5
   SmartTags("D_BarR") = -5

VB script "SetS2"
   SmartTags("D_State") = 2
   SmartTags("D_Bool") = True
   SmartTags("D_SInt") = 12
   SmartTags("D_Int") = 1234
   SmartTags("D_DInt") = 123456
   SmartTags("D_USInt") = 200
   SmartTags("D_UInt") = 40000
   SmartTags("D_UDInt") = 3000000000
   SmartTags("D_Real") = 3.14159
   SmartTags("D_LReal") = 2.718281828
   SmartTags("D_String") = "Hello World"
   SmartTags("D_DateTime") = DateSerial(2026, 11, 22) + TimeSerial(13, 45, 30)
   SmartTags("D_Pct") = 50
   SmartTags("D_Range") = 25
   SmartTags("D_Bits") = 2
   SmartTags("D_Vis") = True
   SmartTags("D_En") = True
   SmartTags("D_X") = 256
   SmartTags("D_Y") = 192
   SmartTags("D_Max") = 200
   SmartTags("D_Min") = -100
   SmartTags("D_TL") = 5
   SmartTags("D_BarR") = 0

VB script "SetS3"
   SmartTags("D_State") = 3
   SmartTags("D_Bool") = True
   SmartTags("D_SInt") = 127
   SmartTags("D_Int") = 32767
   SmartTags("D_DInt") = 2147483647
   SmartTags("D_USInt") = 255
   SmartTags("D_UInt") = 65535
   SmartTags("D_UDInt") = 4294967295
   SmartTags("D_Real") = 123456.789
   SmartTags("D_LReal") = 1E+300
   SmartTags("D_String") = "Ünïcödé äöüß ÄÖÜ € – long text that is wider than the field 0123456789 ABCDEFGHIJ"
   SmartTags("D_DateTime") = DateSerial(2099, 12, 31) + TimeSerial(23, 59, 59)
   SmartTags("D_Pct") = 100
   SmartTags("D_Range") = 75
   SmartTags("D_Bits") = 4
   SmartTags("D_Vis") = True
   SmartTags("D_En") = False
   SmartTags("D_X") = 682
   SmartTags("D_Y") = 384
   SmartTags("D_Max") = 50
   SmartTags("D_Min") = -50
   SmartTags("D_TL") = 10
   SmartTags("D_BarR") = 5

VB script "SetS4"
   SmartTags("D_State") = 4
   SmartTags("D_Bool") = False
   SmartTags("D_SInt") = -1
   SmartTags("D_Int") = -1
   SmartTags("D_DInt") = 0
   SmartTags("D_USInt") = 1
   SmartTags("D_UInt") = 1
   SmartTags("D_UDInt") = 1
   SmartTags("D_Real") = 0.0005
   SmartTags("D_LReal") = -0.0
   SmartTags("D_String") = "äöü ÄÖÜ ß"
   SmartTags("D_DateTime") = DateSerial(1970, 1, 1) + TimeSerial(0, 0, 0)
   SmartTags("D_Pct") = 150
   SmartTags("D_Range") = 200
   SmartTags("D_Bits") = 9
   SmartTags("D_Vis") = False
   SmartTags("D_En") = True
   SmartTags("D_X") = -20
   SmartTags("D_Y") = 0
   SmartTags("D_Max") = 100
   SmartTags("D_Min") = 0
   SmartTags("D_TL") = 50
   SmartTags("D_BarR") = 2.5
*)

(* ===== HMI "HMI_TP900S" =====
system functions are stored by id; their names below are inferred from use

HMI tags "Default tag table"
   "Hmi_Bool" : Bool, internal
   "Hmi_Int" : Int, internal
   "Hmi_Real" : Real, internal
   "Hmi_String" : WString[254], internal

screen "All_Objects" 800x480
   TextField "TextField_1" at 680,10 size 100x30; Text 'Text'
   GraphicView "GraphicView_1" at 10,80 size 100x60
   IOField "IOField_1" at 130,80 size 100x30
   Button "Button_1" at 250,80 size 100x40; TextOff 'Text'
   SymbolicIOField "SymbolicIOField_1" at 370,80 size 120x30; TextOff '0'; TextOn '1'
   GraphicIOField "GraphicIOField_1" at 510,80 size 60x60
   DateTimeField "DateTimeField_1" at 590,80 size 160x30
   Bar "Bar_1" at 10,160 size 40x120
   Switch "Switch_1" at 70,160 size 120x40; CaptionText 'Switch'; TextOff '0'; TextOn '1'
   SymbolLibrary "SymbolLibrary_1" at 210,160 size 60x60
   Slider "Slider_1" at 290,160 size 60x160; Caption 'SIMATIC'
   Gauge "Gauge_1" at 370,160 size 150x150; CaptionText 'SIMATIC'
   Clock "Clock_1" at 540,160 size 150x150

screen "Ctl_01_AlarmView" 800x480, template "Nav"
   AlarmView "Alarm view_1" at 3,3 size 600x300

screen "Ctl_02_TrendView" 800x480, template "Nav"
   TrendView "Trend view_1" at 3,3 size 600x300

screen "Ctl_03_UserView" 800x480, template "Nav"
   UserView "User view_1" at 3,3 size 480x240

screen "Ctl_04_HtmlBrowser" 800x480, template "Nav"
   HTMLBrowser "HTML browser_1" at 3,3 size 192x192

screen "Ctl_05_WatchTable" 800x480, template "Nav"
   StatusForce "Watch table_1" at 3,3 size 600x300; ToolTipText 'Text'

screen "Ctl_06_SmartClientView" 800x480, template "Nav"
   SmartClientView "Sm@rtClient view_1" at 3,3 size 320x240

screen "Ctl_07_RecipeView" 800x480, template "Nav"
   RecipeView "Recipe view_1" at 3,3 size 400x330

screen "Ctl_09_SysDiagView" 800x480, template "Nav"
   SysDiagControl "System diagnostics view_1" at 3,3 size 600x300

screen "Ctl_10_MediaPlayer" 800x480, template "Nav"
   MediaPlayer "Media Player_1" at 3,3 size 240x240

screen "Ctl_11_PlcCodeView" 800x480, template "Nav"
   PLCCodeViewer "PLC code view_1" at 3,3 size 600x300

screen "Ctl_12_GraphOverview" 800x480, template "Nav"
   S7GraphOverview "GRAPH overview_1" at 3,3 size 424x72

screen "Ctl_13_ProDiagOverview" 800x480, template "Nav"
   ProDiagOverview "ProDiag overview_1" at 3,3 size 253x72

screen "Ctl_14_CriteriaAnalysisView" 800x480, template "Nav"
   CriteriaAnalysisView "Criteria analysis view_1" at 3,3 size 460x150

screen "Ctl_15_CameraView" 800x480, template "Nav"
   CameraControl "Camera view_1" at 3,3 size 320x240

screen "Ctl_16_PdfView" 800x480, template "Nav"
   PDFView "PDFView_1" at 3,3 size 320x240

Template "Nav" 800x480
   Button "Nav_01" at 770,2 size 28x22; TextOff 'Text'
      on Click: ActivateScreen("Ctl_01_AlarmView", 0)
   Button "Nav_02" at 770,28 size 28x22; TextOff 'Text'
      on Click: ActivateScreen("Ctl_02_TrendView", 0)
   Button "Nav_03" at 770,54 size 28x22; TextOff 'Text'
      on Click: ActivateScreen("Ctl_03_UserView", 0)
   Button "Nav_04" at 770,80 size 28x22; TextOff 'Text'
      on Click: ActivateScreen("Ctl_04_HtmlBrowser", 0)
   Button "Nav_05" at 770,106 size 28x22; TextOff 'Text'
      on Click: ActivateScreen("Ctl_05_WatchTable", 0)
   Button "Nav_06" at 770,132 size 28x22; TextOff 'Text'
      on Click: ActivateScreen("Ctl_06_SmartClientView", 0)
   Button "Nav_07" at 770,158 size 28x22; TextOff 'Text'
      on Click: ActivateScreen("Ctl_07_RecipeView", 0)
   Button "Nav_09" at 770,210 size 28x22; TextOff 'Text'
      on Click: ActivateScreen("Ctl_09_SysDiagView", 0)
   Button "Nav_10" at 770,236 size 28x22; TextOff 'Text'
      on Click: ActivateScreen("Ctl_10_MediaPlayer", 0)
   Button "Nav_11" at 770,262 size 28x22; TextOff 'Text'
      on Click: ActivateScreen("Ctl_11_PlcCodeView", 0)
   Button "Nav_12" at 770,288 size 28x22; TextOff 'Text'
      on Click: ActivateScreen("Ctl_12_GraphOverview", 0)
   Button "Nav_13" at 770,314 size 28x22; TextOff 'Text'
      on Click: ActivateScreen("Ctl_13_ProDiagOverview", 0)
   Button "Nav_14" at 770,340 size 28x22; TextOff 'Text'
      on Click: ActivateScreen("Ctl_14_CriteriaAnalysisView", 0)
   Button "Nav_15" at 770,366 size 28x22; TextOff 'Text'
      on Click: ActivateScreen("Ctl_15_CameraView", 0)
   Button "Nav_16" at 770,392 size 28x22; TextOff 'Text'
      on Click: ActivateScreen("Ctl_16_PdfView", 0)
   Button "Nav_17" at 770,418 size 28x22; TextOff 'Text'
      on Click: ActivateScreen("All_Objects", 0)
*)

(* ===== HMI "HMI_TP1200" =====
system functions are stored by id; their names below are inferred from use
connection "HMI_Connection_4": ETHERNET, S7_1500_OMS

HMI tags "Default tag table"
   "Hmi_Bool" : Bool, internal
   "Hmi_Int" : Int, internal
   "Hmi_Real" : Real, internal
   "Hmi_String" : WString[254], internal
   "Ext_Bool" : Bool = PLC Plc_Bool AT %M100.0, 1 s
   "Ext_Int" : Int = PLC Plc_Int AT %MW102, 1 s
   "Ext_Real" : Real = PLC Plc_Real AT %MD104, 1 s
   "Ext_Byte" : Byte = PLC Plc_Byte AT %MB108, 1 s

HMI tags "C03_Tags"
   "D_State" : Int, internal
   "D_Bool" : Bool, internal
   "D_SInt" : SInt, internal
   "D_Int" : Int, internal
   "D_DInt" : DInt, internal
   "D_USInt" : USInt, internal
   "D_UInt" : UInt, internal
   "D_UDInt" : UDInt, internal
   "D_Real" : Real, internal
   "D_LReal" : LReal, internal
   "D_String" : WString[254], internal
   "D_DateTime" : DateTime, internal
   "D_Pct" : Int, internal
   "D_Range" : Int, internal
   "D_Bits" : Int, internal
   "D_Vis" : Bool, internal
   "D_En" : Bool, internal
   "D_X" : Int, internal
   "D_Y" : Int, internal
   "D_Max" : Real, internal
   "D_Min" : Real, internal
   "D_TL" : Int, internal
   "D_BarR" : Real, internal

text list "TL_Bit": 0 'Off (0)'; 1 'On (1)'

text list "TL_BitNo": 0 'Bit 0 set'; 1 'Bit 1 set'; 2 'Bit 2 set'; 3 'Bit 3 set'

text list "TL_Value": -100..-1 'Negative (-100..-1)'; 0 'Zero'; 1..9 'One to nine'; 10 'Ten: Ünïcödé äöüß ÄÖÜ €'; 32000 'Undefined value (default entry)'

screen "All_Objects" 1280x800
   TextField "TextField_1" at 680,10 size 100x30; Text 'Text'
   GraphicView "GraphicView_1" at 800,10 size 100x60
   IOField "IOField_1" at 920,10 size 100x30
   Button "Button_1" at 1040,10 size 100x40; TextOff 'Text'
   SymbolicIOField "SymbolicIOField_1" at 10,90 size 120x30; TextOff '0'; TextOn '1'
   GraphicIOField "GraphicIOField_1" at 150,90 size 60x60
   DateTimeField "DateTimeField_1" at 230,90 size 160x30
   Bar "Bar_1" at 410,90 size 40x120
   Switch "Switch_1" at 470,90 size 120x40; CaptionText 'Switch'; TextOff '0'; TextOn '1'
   SymbolLibrary "SymbolLibrary_1" at 610,90 size 60x60
   Slider "Slider_1" at 690,90 size 60x160; Caption 'SIMATIC'
   Gauge "Gauge_1" at 770,90 size 150x150; CaptionText 'SIMATIC'
   Clock "Clock_1" at 940,90 size 150x150

screen "Ctl_01_AlarmView" 1280x800, template "Nav"
   AlarmView "Alarm view_1" at 3,3 size 600x300

screen "Ctl_02_TrendView" 1280x800, template "Nav"
   TrendView "Trend view_1" at 3,3 size 600x300

screen "Ctl_03_UserView" 1280x800, template "Nav"
   UserView "User view_1" at 3,3 size 480x240

screen "Ctl_04_HtmlBrowser" 1280x800, template "Nav"
   HTMLBrowser "HTML browser_1" at 3,3 size 192x192

screen "Ctl_05_WatchTable" 1280x800, template "Nav"
   StatusForce "Watch table_1" at 3,3 size 600x300; ToolTipText 'Text'

screen "Ctl_06_SmartClientView" 1280x800, template "Nav"
   SmartClientView "Sm@rtClient view_1" at 3,3 size 320x240

screen "Ctl_07_RecipeView" 1280x800, template "Nav"
   RecipeView "Recipe view_1" at 3,3 size 400x330

screen "Ctl_09_SysDiagView" 1280x800, template "Nav"
   SysDiagControl "System diagnostics view_1" at 3,3 size 600x300

screen "Ctl_10_MediaPlayer" 1280x800, template "Nav"
   MediaPlayer "Media Player_1" at 3,3 size 240x240

screen "Ctl_15_CameraView" 1280x800, template "Nav"
   CameraControl "Camera view_1" at 3,3 size 320x240

screen "Ctl_16_PdfView" 1280x800, template "Nav"
   PDFView "PDFView_1" at 3,3 size 320x240

Template "Nav" 1280x800
   Button "Nav_01" at 1250,2 size 28x22; TextOff 'Text'
      on Click: ActivateScreen("Ctl_01_AlarmView", 0)
   Button "Nav_02" at 1250,28 size 28x22; TextOff 'Text'
      on Click: ActivateScreen("Ctl_02_TrendView", 0)
   Button "Nav_03" at 1250,54 size 28x22; TextOff 'Text'
      on Click: ActivateScreen("Ctl_03_UserView", 0)
   Button "Nav_04" at 1250,80 size 28x22; TextOff 'Text'
      on Click: ActivateScreen("Ctl_04_HtmlBrowser", 0)
   Button "Nav_05" at 1250,106 size 28x22; TextOff 'Text'
      on Click: ActivateScreen("Ctl_05_WatchTable", 0)
   Button "Nav_06" at 1250,132 size 28x22; TextOff 'Text'
      on Click: ActivateScreen("Ctl_06_SmartClientView", 0)
   Button "Nav_07" at 1250,158 size 28x22; TextOff 'Text'
      on Click: ActivateScreen("Ctl_07_RecipeView", 0)
   Button "Nav_09" at 1250,210 size 28x22; TextOff 'Text'
      on Click: ActivateScreen("Ctl_09_SysDiagView", 0)
   Button "Nav_10" at 1250,236 size 28x22; TextOff 'Text'
      on Click: ActivateScreen("Ctl_10_MediaPlayer", 0)
   Button "Nav_15" at 1250,366 size 28x22; TextOff 'Text'
      on Click: ActivateScreen("Ctl_15_CameraView", 0)
   Button "Nav_16" at 1250,392 size 28x22; TextOff 'Text'
      on Click: ActivateScreen("Ctl_16_PdfView", 0)
   Button "Nav_17" at 1250,418 size 28x22; TextOff 'Text'
      on Click: ActivateScreen("All_Objects", 0)

screen "P_Line_1" 1280x800
   TextField "Label_Default" at 10,62 size 108x16; Text 'Default'
   TextField "Label_BackColor" at 120,62 size 108x16; Text 'BackColor'
   TextField "Label_Color" at 230,62 size 108x16; Text 'Color'
   TextField "Label_EndStyle" at 340,62 size 108x16; Text 'EndStyle'
   TextField "Label_EndStyle_2" at 450,62 size 108x16; Text 'EndStyle_2'
   TextField "Label_EndStyle_3" at 560,62 size 108x16; Text 'EndStyle_3'
   TextField "Label_EndStyle_4" at 670,62 size 108x16; Text 'EndStyle_4'
   TextField "Label_EndStyle_5" at 780,62 size 108x16; Text 'EndStyle_5'
   TextField "Label_FillStyle" at 890,62 size 108x16; Text 'FillStyle'
   TextField "Label_Flashing" at 1000,62 size 108x16; Text 'Flashing'
   TextField "Label_LineEndShapeStyle_2" at 1110,62 size 108x16; Text 'LineEndShapeStyle_2'
   TextField "Label_LineWidth" at 10,138 size 108x16; Text 'LineWidth'
   TextField "Label_StartStyle" at 120,138 size 108x16; Text 'StartStyle'
   TextField "Label_StartStyle_2" at 230,138 size 108x16; Text 'StartStyle_2'
   TextField "Label_StartStyle_3" at 340,138 size 108x16; Text 'StartStyle_3'
   TextField "Label_StartStyle_4" at 450,138 size 108x16; Text 'StartStyle_4'
   TextField "Label_StartStyle_5" at 560,138 size 108x16; Text 'StartStyle_5'
   TextField "Label_Style" at 670,138 size 108x16; Text 'Style'
   TextField "Label_Style_2" at 780,138 size 108x16; Text 'Style_2'
   TextField "Label_Style_3" at 890,138 size 108x16; Text 'Style_3'
   TextField "Label_Style_4" at 1000,138 size 108x16; Text 'Style_4'
   TextField "Label_UseDesignColorSchema" at 1110,138 size 108x16; Text 'UseDesignColorSchema'
   Button "Next" at 1238,776 size 40x22; TextOff 'Text'
      on Click: ActivateScreen("P_Polyline_1", 0)

screen "P_Polyline_1" 1280x800
   TextField "Label_Default" at 10,62 size 108x16; Text 'Default'
   TextField "Label_BackColor" at 120,62 size 108x16; Text 'BackColor'
   TextField "Label_Color" at 230,62 size 108x16; Text 'Color'
   TextField "Label_EndStyle" at 340,62 size 108x16; Text 'EndStyle'
   TextField "Label_EndStyle_2" at 450,62 size 108x16; Text 'EndStyle_2'
   TextField "Label_EndStyle_3" at 560,62 size 108x16; Text 'EndStyle_3'
   TextField "Label_EndStyle_4" at 670,62 size 108x16; Text 'EndStyle_4'
   TextField "Label_EndStyle_5" at 780,62 size 108x16; Text 'EndStyle_5'
   TextField "Label_FillStyle" at 890,62 size 108x16; Text 'FillStyle'
   TextField "Label_Flashing" at 1000,62 size 108x16; Text 'Flashing'
   TextField "Label_LineEndShapeStyle_2" at 1110,62 size 108x16; Text 'LineEndShapeStyle_2'
   TextField "Label_LineWidth" at 10,138 size 108x16; Text 'LineWidth'
   TextField "Label_StartStyle" at 120,138 size 108x16; Text 'StartStyle'
   TextField "Label_StartStyle_2" at 230,138 size 108x16; Text 'StartStyle_2'
   TextField "Label_StartStyle_3" at 340,138 size 108x16; Text 'StartStyle_3'
   TextField "Label_StartStyle_4" at 450,138 size 108x16; Text 'StartStyle_4'
   TextField "Label_StartStyle_5" at 560,138 size 108x16; Text 'StartStyle_5'
   TextField "Label_Style" at 670,138 size 108x16; Text 'Style'
   TextField "Label_Style_2" at 780,138 size 108x16; Text 'Style_2'
   TextField "Label_Style_3" at 890,138 size 108x16; Text 'Style_3'
   TextField "Label_Style_4" at 1000,138 size 108x16; Text 'Style_4'
   TextField "Label_UseDesignColorSchema" at 1110,138 size 108x16; Text 'UseDesignColorSchema'
   Button "Next" at 1238,776 size 40x22; TextOff 'Text'
      on Click: ActivateScreen("P_Polygon_1", 0)

screen "P_Polygon_1" 1280x800
   TextField "Label_Default" at 10,62 size 108x16; Text 'Default'
   TextField "Label_BackColor" at 120,62 size 108x16; Text 'BackColor'
   TextField "Label_BackFillStyle" at 230,62 size 108x16; Text 'BackFillStyle'
   TextField "Label_BorderColor" at 340,62 size 108x16; Text 'BorderColor'
   TextField "Label_BorderWidth" at 450,62 size 108x16; Text 'BorderWidth'
   TextField "Label_EdgeStyle" at 560,62 size 108x16; Text 'EdgeStyle'
   TextField "Label_EdgeStyle_2" at 670,62 size 108x16; Text 'EdgeStyle_2'
   TextField "Label_EdgeStyle_3" at 780,62 size 108x16; Text 'EdgeStyle_3'
   TextField "Label_EdgeStyle_4" at 890,62 size 108x16; Text 'EdgeStyle_4'
   TextField "Label_Flashing" at 1000,62 size 108x16; Text 'Flashing'
   TextField "Label_UseDesignColorSchema" at 1110,62 size 108x16; Text 'UseDesignColorSchema'
   Button "Next" at 1238,776 size 40x22; TextOff 'Text'
      on Click: ActivateScreen("P_Ellipse_1", 0)

screen "P_Ellipse_1" 1280x800
   TextField "Label_Default" at 10,62 size 108x16; Text 'Default'
   TextField "Label_BackColor" at 120,62 size 108x16; Text 'BackColor'
   TextField "Label_BackFillStyle" at 230,62 size 108x16; Text 'BackFillStyle'
   TextField "Label_BorderColor" at 340,62 size 108x16; Text 'BorderColor'
   TextField "Label_BorderWidth" at 450,62 size 108x16; Text 'BorderWidth'
   TextField "Label_EdgeStyle" at 560,62 size 108x16; Text 'EdgeStyle'
   TextField "Label_EdgeStyle_2" at 670,62 size 108x16; Text 'EdgeStyle_2'
   TextField "Label_EdgeStyle_3" at 780,62 size 108x16; Text 'EdgeStyle_3'
   TextField "Label_EdgeStyle_4" at 890,62 size 108x16; Text 'EdgeStyle_4'
   TextField "Label_Flashing" at 1000,62 size 108x16; Text 'Flashing'
   TextField "Label_UseDesignColorSchema" at 1110,62 size 108x16; Text 'UseDesignColorSchema'
   Button "Next" at 1238,776 size 40x22; TextOff 'Text'
      on Click: ActivateScreen("P_Circle_1", 0)

screen "P_Circle_1" 1280x800
   TextField "Label_Default" at 10,62 size 58x16; Text 'Default'
   TextField "Label_BackColor" at 70,62 size 58x16; Text 'BackColor'
   TextField "Label_BackFillStyle" at 130,62 size 58x16; Text 'BackFillStyle'
   TextField "Label_BorderColor" at 190,62 size 58x16; Text 'BorderColor'
   TextField "Label_BorderWidth" at 250,62 size 58x16; Text 'BorderWidth'
   TextField "Label_EdgeStyle" at 310,62 size 58x16; Text 'EdgeStyle'
   TextField "Label_EdgeStyle_2" at 370,62 size 58x16; Text 'EdgeStyle_2'
   TextField "Label_EdgeStyle_3" at 430,62 size 58x16; Text 'EdgeStyle_3'
   TextField "Label_EdgeStyle_4" at 490,62 size 58x16; Text 'EdgeStyle_4'
   TextField "Label_Flashing" at 550,62 size 58x16; Text 'Flashing'
   TextField "Label_UseDesignColorSchema" at 610,62 size 58x16; Text 'UseDesignColorSchema'
   Button "Next" at 1238,776 size 40x22; TextOff 'Text'
      on Click: ActivateScreen("P_Rectangle_1", 0)

screen "P_Rectangle_1" 1280x800
   TextField "Label_Default" at 10,62 size 108x16; Text 'Default'
   TextField "Label_BackColor" at 120,62 size 108x16; Text 'BackColor'
   TextField "Label_BackFillStyle" at 230,62 size 108x16; Text 'BackFillStyle'
   TextField "Label_BorderColor" at 340,62 size 108x16; Text 'BorderColor'
   TextField "Label_BorderWidth" at 450,62 size 108x16; Text 'BorderWidth'
   TextField "Label_EdgeStyle" at 560,62 size 108x16; Text 'EdgeStyle'
   TextField "Label_EdgeStyle_2" at 670,62 size 108x16; Text 'EdgeStyle_2'
   TextField "Label_EdgeStyle_3" at 780,62 size 108x16; Text 'EdgeStyle_3'
   TextField "Label_EdgeStyle_4" at 890,62 size 108x16; Text 'EdgeStyle_4'
   TextField "Label_Flashing" at 1000,62 size 108x16; Text 'Flashing'
   TextField "Label_RoundCornerHeight" at 1110,62 size 108x16; Text 'RoundCornerHeight'
   TextField "Label_RoundCornerWidth" at 10,138 size 108x16; Text 'RoundCornerWidth'
   TextField "Label_UseDesignColorSchema" at 120,138 size 108x16; Text 'UseDesignColorSchema'
   Button "Next" at 1238,776 size 40x22; TextOff 'Text'
      on Click: ActivateScreen("P_TextField_1", 0)

screen "P_TextField_1" 1280x800
   TextField "Default" at 10,10 size 100x30; Text 'Text'
   TextField "Label_Default" at 10,42 size 108x16; Text 'Default'
   TextField "BackColor" at 120,10 size 100x30; Text 'Text'
   TextField "Label_BackColor" at 120,42 size 108x16; Text 'BackColor'
   TextField "BackFillStyle" at 230,10 size 100x30; Text 'Text'
   TextField "Label_BackFillStyle" at 230,42 size 108x16; Text 'BackFillStyle'
   TextField "BorderBackColor" at 340,10 size 100x30; Text 'Text'
   TextField "Label_BorderBackColor" at 340,42 size 108x16; Text 'BorderBackColor'
   TextField "BorderColor" at 450,10 size 100x30; Text 'Text'
   TextField "Label_BorderColor" at 450,42 size 108x16; Text 'BorderColor'
   TextField "BorderWidth" at 560,10 size 100x30; Text 'Text'
   TextField "Label_BorderWidth" at 560,42 size 108x16; Text 'BorderWidth'
   TextField "BottomMargin" at 670,10 size 100x30; Text 'Text'
   TextField "Label_BottomMargin" at 670,42 size 108x16; Text 'BottomMargin'
   TextField "CornerRadius" at 780,10 size 100x30; Text 'Text'
   TextField "Label_CornerRadius" at 780,42 size 108x16; Text 'CornerRadius'
   TextField "EdgeStyle" at 890,10 size 100x30; Text 'Text'
   TextField "Label_EdgeStyle" at 890,42 size 108x16; Text 'EdgeStyle'
   TextField "EdgeStyle_2" at 1000,10 size 100x30; Text 'Text'
   TextField "Label_EdgeStyle_2" at 1000,42 size 108x16; Text 'EdgeStyle_2'
   TextField "EdgeStyle_3" at 1110,10 size 100x30; Text 'Text'
   TextField "Label_EdgeStyle_3" at 1110,42 size 108x16; Text 'EdgeStyle_3'
   TextField "EdgeStyle_4" at 10,66 size 100x30; Text 'Text'
   TextField "Label_EdgeStyle_4" at 10,98 size 108x16; Text 'EdgeStyle_4'
   TextField "FitToLargest" at 120,66 size 100x30; Text 'Text'
   TextField "Label_FitToLargest" at 120,98 size 108x16; Text 'FitToLargest'
   TextField "Flashing" at 230,66 size 100x30; Text 'Text'
   TextField "Label_Flashing" at 230,98 size 108x16; Text 'Flashing'
   TextField "ForeColor" at 340,66 size 100x30; Text 'Text'
   TextField "Label_ForeColor" at 340,98 size 108x16; Text 'ForeColor'
   TextField "HorizontalAlignment" at 450,66 size 100x30; Text 'Text'
   TextField "Label_HorizontalAlignment" at 450,98 size 108x16; Text 'HorizontalAlignment'
   TextField "HorizontalAlignment_2" at 560,66 size 100x30; Text 'Text'
   TextField "Label_HorizontalAlignment_2" at 560,98 size 108x16; Text 'HorizontalAlignment_2'
   TextField "LeftMargin" at 670,66 size 100x30; Text 'Text'
   TextField "Label_LeftMargin" at 670,98 size 108x16; Text 'LeftMargin'
   TextField "RightMargin" at 780,66 size 100x30; Text 'Text'
   TextField "Label_RightMargin" at 780,98 size 108x16; Text 'RightMargin'
   TextField "TopMargin" at 890,66 size 100x30; Text 'Text'
   TextField "Label_TopMargin" at 890,98 size 108x16; Text 'TopMargin'
   TextField "UseDesignColorSchema" at 1000,66 size 100x30; Text 'Text'
   TextField "Label_UseDesignColorSchema" at 1000,98 size 108x16; Text 'UseDesignColorSchema'
   TextField "VerticalAlignment" at 1110,66 size 100x30; Text 'Text'
   TextField "Label_VerticalAlignment" at 1110,98 size 108x16; Text 'VerticalAlignment'
   TextField "VerticalAlignment_2" at 10,122 size 100x30; Text 'Text'
   TextField "Label_VerticalAlignment_2" at 10,154 size 108x16; Text 'VerticalAlignment_2'
   Button "Next" at 1238,776 size 40x22; TextOff 'Text'
      on Click: ActivateScreen("P_GraphicView_1", 0)

